(* IEC 61131-3 sources: daoli-st-library/DL_Algo, 207 files *)

(* ---- FB_DL_AdaptiveLeadLag.st ---- *)
(*==============================================================================
 * 组件名称 (Component)  : FB_DL_AdaptiveLeadLag
 * 所属子库 (Sublibrary) : DL_Algo
 * 当前版本 (Version)    : 1.0.0
 * 兼容性   (Platform)   : CODESYS 3.5+ / TwinCAT 3 / 汇川 InoProShop / 施耐德 Machine Expert
 *                         仅依赖 Standard.library（R_TRIG / ABS），零厂商私有库
 * 功能描述 (Function)   : 自适应超前-滞后补偿（误差驱动参数缓调 + 无扰切换）。
 *                         ① 补偿本体：连续式 G(s) = (1 + Tlead·s) / (1 + Tlag·s) 的离散实现
 *                            超前段：yLead = x + Tlead·(x − xPrev) / fDtS
 *                            滞后段：y     = y + (yLead − y) · fDtS / (Tlag + fDtS)
 *                            两段都用 fDtS（调用方给的采样周期，秒），**不做 TIME→数值转换**。
 *                         ② 参数缓调：Tlead 按误差幅值缓升缓降（相位裕度需求随误差增大），
 *                            每拍步长 = fAdaptGain·|fErr|·fDtS，并被 fAdaptRate·fDtS 限幅
 *                            （限幅保证"缓"：参数变化速度受控，不会一拍跳变引起输出突跳）。
 *                            Tlead 始终钳在 [fTleadMin, fTleadMax]。
 *                         ③ 无扰切换：bEnable 上升沿开始，fBlend 以固定步长 fDtS / fRampSec
 *                            从 0 线性升到 1；输出 = 切换前保持值 + blend·(计算值 − 保持值)。
 *                            **不用 TON 的 ET 做斜坡**，因而无 TIME→数值转换（跨平台一致），
 *                            且斜坡长度由 fRampSec 显式给出，可预测、可复现。
 * 接口     (Interface)  : 输入 fIn 输入信号、fErr 跟踪误差（驱动自适应）、fDtS 采样周期（秒）、
 *                         fTleadInit / fTlagInit 初值、fTleadMin / fTleadMax 超前时间限、
 *                         fAdaptGain 自适应增益、fAdaptRate 参数变化率限、fRampSec 无扰斜坡时长、
 *                         fOutMax 输出饱和限、bEnable 使能、bReset 复位；输出 fOut 补偿输出、
 *                         fTleadUsed / fTlagUsed 实际使用参数、fBlend 切换斜坡进度、bActive 已生效、
 *                         bLimited 输出饱和、eState / eCause / bError。
 * 边界     (Boundary)   : ① **属主边界（写死）：本件是补偿器本体，输出 fOut 供上层注入，
 *                         不直接写轴指令/不进闭环回路**；本件不做参数辨识（辨识属 `FB_DL_RlsEstimator`），
 *                         只按误差缓调。
 *                         ② 组态闸：fDtS <= DL_ALL_EPS（除零 + 步长退化）、fTlagInit < 0.0、
 *                         fTleadMin < 0.0、fTleadMax <= fTleadMin、fAdaptGain < 0.0、
 *                         fAdaptRate <= 0.0、fRampSec <= DL_ALL_EPS、fOutMax <= 0.0、任一 NaN
 *                         → 故障锁存，fOut 置 0（安全侧）。
 *                         ③ bEnable=FALSE 语义（R191 声明）：fOut 立即置 0（补偿器禁用即不注入），
 *                         但**保留 fTleadUsed 与内部滞后状态**，下次使能由 fBlend 斜坡重新接续，
 *                         属"冻结参数、清零输出"，与"复位"（参数回初值）不同。
 *                         ④ 单枚 R_TRIG（bReset 与 bEnable 各一枚）段 0 无条件周期刷新。
 *                         ⑤ 故障相迁出唯一路径 = bReset 上升沿（R228B）。
 *                         ⑥ 零全局耦合（无 GVL / 无 VAR_EXTERNAL / 无物理地址）。
 * 分工声明 (Scope)      : 与 `FB_DL_StribeckFrictionComp`（摩擦模型本体）分工——本件是线性
 *                         超前滞后相位补偿，那件是非线性摩擦补偿；两者可并行相加注入，
 *                         但都不自己注入（注入点唯一）。
 * 来源标签 (Source Tag) : T2-1 ◐（公开经典超前-滞后补偿结构与自适应步长思想，参考参数域，
 *                         零代码行复制；固定步长无扰斜坡为本库自研包装）
 * 解除式   (Release)    : bReset 上升沿 ∧ 组态合法 → 清故障、参数回初值、清滞后状态与斜坡。
 *                         自证可满足：复位不依赖锁存量。
 * 码表     (Codes)      : 本件不占用任何全局数字码位。出口为 REAL + BOOL（bActive / bLimited /
 *                         bError）+ ENUM（eState / eCause）；数字码位待主控收口阶段统一派号。
 * 红线自检 (Redline)    : R1 ✓ 零 GVL/VAR_EXTERNAL ｜ R2 ✓ 零 %I/%Q/%M ｜ R3 ✓ 纯 IEC 61131-3
 *                         R4 ✓ 除零闸 + 参数区间闸 + 输出饱和 + NaN 闸 ｜ R5 ✓ 声明逐行同行双语注释
 *                         R6 ✓ ENUM+CASE 含 ELSE ｜ R7 ✓ R_TRIG 段 0 无条件刷新
 * 修订历史 (Revision)   : 2026-11-19  v1.0.0  R46 首版（批次 4 · 序号 17）
 *==============================================================================*)

TYPE E_DL_AllState :
(
    eIdle  := 0,    // 未使能或未完成切换斜坡 / Disabled, ramp not started
    eRamp  := 10,   // 无扰切换斜坡进行中 / Bumpless transfer ramp in progress
    eRun   := 20,   // 补偿器全效运行 / Compensator fully engaged
    eFault := 90    // 组态故障相 / Configuration fault phase
);
END_TYPE

TYPE E_DL_AllCause :
(
    eNone       := 0,   // 无异常 / No anomaly
    eCfgIllegal := 1,   // 组态非法（采样周期/时间限/增益/非有限） / Illegal configuration
    eOutSat     := 2,   // 输出触饱和（补偿量需求超限） / Output saturated
    ePhaseBad   := 3    // 非法相位兜底 / Illegal phase fallback
);
END_TYPE

FUNCTION_BLOCK FB_DL_AdaptiveLeadLag
VAR_INPUT
    fIn        : REAL := 0.0;       // 输入信号 [工程单位] / Input signal [unit]
    fErr       : REAL := 0.0;       // 跟踪误差（驱动自适应） [工程单位] / Tracking error driving the adaptation [unit]
    fDtS       : REAL := 0.001;     // 采样周期，域 > DL_ALL_EPS [s] / Sample period, domain > epsilon [s]
    fTleadInit : REAL := 0.05;      // 超前时间初值，域 >= 0.0 [s] / Initial lead time, >= 0.0 [s]
    fTlagInit  : REAL := 0.20;      // 滞后时间初值，域 >= 0.0 [s] / Initial lag time, >= 0.0 [s]
    fTleadMin  : REAL := 0.01;      // 超前时间下限，域 >= 0.0 [s] / Lead time lower bound, >= 0.0 [s]
    fTleadMax  : REAL := 0.50;      // 超前时间上限，域 > fTleadMin [s] / Lead time upper bound, > lower [s]
    fAdaptGain : REAL := 0.10;      // 自适应增益，域 >= 0.0 [1/s] / Adaptation gain, >= 0.0 [1/s]
    fAdaptRate : REAL := 0.50;      // 参数变化率限，域 > 0.0 [s/s] / Parameter rate limit, > 0.0 [s/s]
    fRampSec   : REAL := 0.20;      // 无扰斜坡时长，域 > DL_ALL_EPS [s] / Bumpless ramp duration, > epsilon [s]
    fOutMax    : REAL := 100.0;     // 输出饱和限，域 > 0.0 [工程单位] / Output saturation limit, > 0.0 [unit]
    bEnable    : BOOL := FALSE;     // 使能；FALSE 时输出置 0 但保留参数 [-] / Enable; FALSE zeroes the output but keeps parameters
    bReset     : BOOL := FALSE;     // 复位，上升沿清故障并使参数回初值 [-] / Reset, clears the fault and restores initial parameters
END_VAR
VAR_OUTPUT
    fOut       : REAL;              // 补偿输出（已饱和） [工程单位] / Compensation output, saturated [unit]
    fTleadUsed : REAL;              // 实际使用中的超前时间 [s] / Lead time in use [s]
    fTlagUsed  : REAL;              // 实际使用中的滞后时间 [s] / Lag time in use [s]
    fBlend     : REAL;              // 切换斜坡进度，域 0..1 [-] / Ramp progress in 0..1
    bActive    : BOOL;              // 补偿器全效生效（blend 已达 1） [-] / Compensator fully engaged
    bLimited   : BOOL;              // 本拍输出触饱和 [-] / Output saturated this scan
    eState     : E_DL_AllState;     // 状态出口 [-] / State outlet
    eCause     : E_DL_AllCause;     // 成因出口（R190 归因唯一） [-] / Cause outlet
    bError     : BOOL;              // 故障标志（组态非法） [-] / Error flag, illegal configuration
END_VAR
VAR
    _eState  : E_DL_AllState := E_DL_AllState.eIdle;    // 内部相位（CASE 唯一写入目标） / Internal phase
    _eCause  : E_DL_AllCause := E_DL_AllCause.eNone;    // 成因出口暂存 / Cause staging
    rtReset  : R_TRIG;              // 复位沿实例，段 0 无条件调用 / Reset edge instance
    rtEnable : R_TRIG;              // 使能沿实例，段 0 无条件调用 / Enable edge instance
    _fTlead  : REAL;                // 超前时间（锁存量） [s] / Lead time, latched [s]
    _fXPrev  : REAL;                // 上拍输入快照（锁存量） [工程单位] / Previous input, latched [unit]
    _fYState : REAL;                // 滞后段内部状态（锁存量） [工程单位] / Lag stage internal state, latched [unit]
    _fBlend  : REAL;                // 斜坡进度（锁存量） [-] / Ramp progress, latched
    _fHold   : REAL;                // 切换前保持值（锁存量） [工程单位] / Value held before transfer, latched [unit]
    _fLead   : REAL;                // 超前段输出当拍量 [工程单位] / Lead-stage output this scan [unit]
    _fComp   : REAL;                // 补偿计算值当拍量 [工程单位] / Computed compensation this scan [unit]
    _fStep   : REAL;                // 参数调整步长当拍量 [s] / Parameter step this scan [s]
    _fRate   : REAL;                // 每拍允许的最大参数变化量 [s] / Maximum parameter change per scan [s]
    _bFault  : BOOL;                // 组态故障锁存位（锁存量） / Latched configuration fault
    _bCfgBad : BOOL;                // 组态非法当拍量 [-] / Illegal configuration this scan
    _bNonFin : BOOL;                // 输入非有限当拍量 [-] / Non-finite input this scan
    _bSat    : BOOL;                // 本拍输出饱和当拍量 [-] / Output saturation this scan
END_VAR
VAR CONSTANT
    DL_ALL_EPS  : REAL := 1.0E-9;   // 时间判零容差（秒级，需比通用 eps 更紧） [无量纲] / Time epsilon in seconds, tighter than usual
    DL_ALL_ONE  : REAL := 1.0;      // 斜坡进度上限 1.0 [无量纲] / Ramp ceiling
    DL_ALL_ZERO : REAL := 0.0;      // 零基准 [无量纲] / Zero baseline
END_VAR

(* —— 段 0：判据派生 + 两沿实例无条件周期刷新 —— *)
_bNonFin := (fIn <> fIn) OR (fErr <> fErr) OR (fDtS <> fDtS)              // NaN 自反判（判等禁令唯一例外） / NaN self-reflexive tests
         OR (fTleadInit <> fTleadInit) OR (fTlagInit <> fTlagInit)
         OR (fTleadMin <> fTleadMin) OR (fTleadMax <> fTleadMax)
         OR (fAdaptGain <> fAdaptGain) OR (fAdaptRate <> fAdaptRate)
         OR (fRampSec <> fRampSec) OR (fOutMax <> fOutMax);
_bCfgBad := (fDtS <= DL_ALL_EPS)                                          // 采样周期闸（除零 + 步长退化） / Sample period gate
         OR (fTleadInit < 0.0) OR (fTlagInit < 0.0)                       // 时间初值非负闸 / Non-negative initial times
         OR (fTleadMin < 0.0) OR (fTleadMax <= fTleadMin)                 // 超前限区间闸 / Lead bounds interval gate
         OR (fAdaptGain < 0.0) OR (fAdaptRate <= 0.0)                     // 自适应增益与速率闸 / Adaptation gain and rate gates
         OR (fRampSec <= DL_ALL_EPS) OR (fOutMax <= 0.0) OR _bNonFin;     // 斜坡与饱和限 + 非有限 / Ramp, saturation limit, non-finite
rtReset(CLK := bReset);                                                   // 复位沿，每拍必调（R228A） / Reset edge, every scan
rtEnable(CLK := bEnable);                                                 // 使能沿，每拍必调 / Enable edge, every scan

(* —— 段 1：单拍量预清零（锁存量 _fTlead/_fXPrev/_fYState/_fBlend/_fHold/_bFault 不入清单） —— *)
fOut     := 0.0;        // 输出每拍预清 / Output preset
fBlend   := 0.0;        // 斜坡出口预清 / Ramp outlet preset
bActive  := FALSE;      // 生效位预清 / Active preset
bLimited := FALSE;      // 饱和位预清 / Limited preset
bError   := FALSE;      // 故障标志预清（R45 配对） / Error flag preset
_bSat    := FALSE;      // 饱和当拍量预清 / Saturation preset

(* —— 段 2：复位沿（参数回初值、清滞后状态与斜坡） —— *)
IF rtReset.Q THEN
    _bFault  := FALSE;                       // 清故障锁存 / Clear the fault latch
    _eCause  := E_DL_AllCause.eNone;         // 清成因 / Clear cause
    _fTlead  := fTleadInit;                  // 超前时间回初值 / Lead time back to the initial value
    _fYState := 0.0;                         // 滞后段状态清零 / Lag state cleared
    _fXPrev  := fIn;                         // 输入快照对齐当拍（防复位首拍伪微分） / Align the snapshot to the present input
    _fBlend  := 0.0;                         // 斜坡清零 / Ramp cleared
    _fHold   := 0.0;                         // 保持值清零 / Hold cleared
    IF _eState = E_DL_AllState.eFault THEN
        _eState := E_DL_AllState.eIdle;      // 故障相迁出（R228B） / Leave fault phase
    END_IF
END_IF
IF _bCfgBad THEN
    _bFault := TRUE;                         // 组态非法锁存 / Latch illegal configuration
    _eCause := E_DL_AllCause.eCfgIllegal;    // 归因：组态非法 / Cause: illegal configuration
END_IF

(* —— 段 3：无扰切换斜坡管理（使能沿起坡；固定步长，无 TIME→数值转换） —— *)
IF rtEnable.Q THEN
    _fHold  := fOut;                         // 记录切换前输出为保持值（若无历史则为 0） / Capture the pre-transfer output
    _fBlend := 0.0;                          // 从 0 起坡 / Start the ramp at zero
    _eState := E_DL_AllState.eRamp;          // 入斜坡相 / Enter the ramp phase
END_IF
IF bEnable AND (NOT _bCfgBad) THEN
    IF _fBlend < DL_ALL_ONE THEN
        _fBlend := _fBlend + (fDtS / fRampSec);     // 固定步长推进（分母已闸） / Fixed-step advance, denominator gated
        IF _fBlend >= DL_ALL_ONE THEN
            _fBlend := DL_ALL_ONE;                  // 上限钳 / Ceiling clamp
            _eState := E_DL_AllState.eRun;           // 斜坡完成，全效运行 / Ramp done, fully engaged
        ELSE
            _eState := E_DL_AllState.eRamp;          // 仍在斜坡 / Still ramping
        END_IF
    END_IF
ELSIF NOT bEnable THEN
    _fBlend := 0.0;                                 // 禁用即清坡（下次使能重新无扰起坡） / Disable clears the ramp
END_IF

(* —— 段 4：自适应参数缓调（误差驱动，速率限幅，区间钳位） —— *)
IF bEnable AND (NOT _bCfgBad) THEN
    _fStep := fAdaptGain * ABS(fErr) * fDtS;                    // 误差驱动的期望步长 [s] / Desired step from the error
    _fRate := fAdaptRate * fDtS;                                // 每拍允许的最大变化量 [s] / Allowed change per scan
    IF _fStep > _fRate THEN
        _fStep := _fRate;                                       // 速率限幅（"缓"调的实现点） / Rate limit, where "slow" is enforced
    END_IF
    IF fErr > 0.0 THEN
        _fTlead := _fTlead + _fStep;                            // 误差为正：加大超前 / Positive error increases the lead
    ELSE
        _fTlead := _fTlead - _fStep;                            // 误差为负：减小超前 / Negative error reduces the lead
    END_IF
    IF _fTlead > fTleadMax THEN
        _fTlead := fTleadMax;                                   // 上限钳 / Upper clamp
    END_IF
    IF _fTlead < fTleadMin THEN
        _fTlead := fTleadMin;                                   // 下限钳 / Lower clamp
    END_IF
END_IF

(* —— 段 5：补偿本体计算（超前段 → 滞后段） —— *)
IF bEnable AND (NOT _bCfgBad) THEN
    _fLead := fIn + (_fTlead * ((fIn - _fXPrev) / fDtS));       // 超前段（分母已闸） / Lead stage, denominator gated
    IF (fTlagInit + fDtS) > DL_ALL_EPS THEN
        _fYState := _fYState + ((_fLead - _fYState) * (fDtS / (fTlagInit + fDtS)));   // 滞后段一阶离散 / Lag stage, first order
    ELSE
        _fYState := _fLead;                                     // 滞后时间为 0 且 dt 病态：直通 / Degenerate case: pass through
    END_IF
    _fComp := _fYState;                                         // 补偿计算值 / Computed compensation
    fOut   := _fHold + (_fBlend * (_fComp - _fHold));           // 无扰混合输出 / Bumpless blended output
    IF fOut > fOutMax THEN
        fOut   := fOutMax;                                      // 正饱和 / Saturate high
        _bSat  := TRUE;
    ELSIF fOut < -fOutMax THEN
        fOut   := -fOutMax;                                     // 负饱和 / Saturate low
        _bSat  := TRUE;
    END_IF
    _fXPrev := fIn;                                             // 输入快照更新（本拍末） / Input snapshot at body end
END_IF

(* —— 段 6：锁存相位迁移闸 —— *)
IF _bFault AND (_eState <> E_DL_AllState.eFault) THEN
    _eState := E_DL_AllState.eFault;                            // 锁存即入故障相 / Latch enters fault phase
END_IF

(* —— 段 7：相位机（ENUM 全成员显式标签 + ELSE 兜底，R128） —— *)
CASE _eState OF

E_DL_AllState.eIdle:
    IF _bFault THEN                                             // 出口 1：组态故障 / Configuration fault
        _eState := E_DL_AllState.eFault;
    ELSIF bEnable THEN                                          // 出口 2：使能到来（无沿也算） / Enable present
        _eState := E_DL_AllState.eRamp;
    END_IF

E_DL_AllState.eRamp:
    IF _bFault THEN                                             // 出口 1：组态故障 / Configuration fault
        _eState := E_DL_AllState.eFault;
    ELSIF (NOT bEnable) THEN                                    // 出口 2：被禁用，回等待相 / Disabled, back to idle
        _eState := E_DL_AllState.eIdle;
    END_IF

E_DL_AllState.eRun:
    IF _bFault THEN                                             // 出口 1：组态故障 / Configuration fault
        _eState := E_DL_AllState.eFault;
    ELSIF NOT bEnable THEN                                      // 出口 2：被禁用，回等待相 / Disabled, back to idle
        _eState := E_DL_AllState.eIdle;
    END_IF

E_DL_AllState.eFault:
    ;                                                           // 故障相：仅段 2 复位沿可迁出 / Only the reset edge leaves this phase

ELSE
    _bFault := TRUE;                                            // 非法相位兜底锁存 / Illegal-phase fallback latch
    _eCause := E_DL_AllCause.ePhaseBad;                         // 归因：非法相位 / Cause: illegal phase
    _eState := E_DL_AllState.eFault;                            // 强拉故障相 / Force fault phase

END_CASE

(* —— 段 8：出口单点映射（名实双出口，R191） —— *)
fTleadUsed := _fTlead;                                          // 超前时间出口 / Lead time outlet
fTlagUsed  := fTlagInit;                                        // 滞后时间出口（本件不调整滞后） / Lag time outlet, not adapted
fBlend     := _fBlend;                                          // 斜坡出口 / Ramp outlet
bActive    := (_eState = E_DL_AllState.eRun) AND (NOT _bFault); // 全效 = 运行相且无故障 / Fully engaged
bLimited   := _bSat;                                            // 饱和出口 / Saturation outlet
bError     := _bFault OR _bCfgBad;                              // 故障标志 = 锁存或组态非法 / Error = latch or illegal config
IF _bSat AND (NOT _bFault) THEN
    _eCause := E_DL_AllCause.eOutSat;                           // 提示：输出饱和（信息级） / Notice: output saturated
END_IF
eState := _eState;                                              // 状态出口 / State outlet
eCause := _eCause;                                              // 成因出口 / Cause outlet

END_FUNCTION_BLOCK

(* ---- FB_DL_CrossLimitSelect.st ---- *)
(*==============================================================================
 * 组件名称 (Component)  : FB_DL_CrossLimitSelect
 * 溯源说明 (Provenance): 道莅 clean-room 防御性实现（IEC 61131-3 纯净实现，闭源文档仅借语义，零代码行）
 * 所属子库 (Sublibrary) : DL_Algo / ProcessControl
 * 当前版本 (Version)    : 1.0.0
 * 兼容性   (Platform)   : CODESYS 3.5 / TwinCAT 3 / 汇川 InoProShop / 施耐德
 *                         Machine Expert；纯 IEC 61131-3（第 3 版），仅用
 *                         Standard.library 的 LIMIT / MIN / MAX / ABS
 * 组件分类 (Category)   : 功能块（FUNCTION_BLOCK）· 燃烧双交叉限幅
 * 功能一句话 (Summary)  : 把主控输出分配成空气/燃气两路给定，按「先行侧自由、
 *                         跟随侧受实测流量约束」的双交叉限幅律钳制，输出限幅
 *                         标志与距限幅点余量。
 *
 * 本件存在的意义 (Why this unit exists)
 *   库内 SplitRangeControl 是单输出分程、RatioController 是比值站，都不解
 *   「空燃两侧谁先给」这个燃烧专有语义。双交叉限幅管的是**同拍的选择律**：
 *   升负荷时先行侧先动、跟随侧被实测流量压住；降负荷时反过来。
 *   写成一件的理由是它必须逐拍可复算（验收向量要能独立手算），
 *   与氧量修正（慢时标积分律，见 FB_DL_ExcessAirTrim）不可合并。
 *
 * 依赖收窄 (Dependency narrowing)
 *   DL_Algo 只允许依赖 Standard.library（DL_Algo/VERSION.md 明示不得引用
 *   DL_Base / DL_MathData）。因此本件的限幅用内建 LIMIT、容差比较与死区
 *   判断全部内联等价实现，不调用任何 DL_ 子库件。此处声明留档（R11 先例）。
 *
 * 折算口径 (Scaling rationale —— 必须写清，否则本件不可复算)
 *   主控输出是 [%]，流量是 [Nm3/h]，两者不同量纲，接口未给阀门流量量程。
 *   本件的折算基准是**实测流量本身**：主控 [%] 与实测流量在当前工况下对应，
 *   故「约束侧的允许百分比」= 主控输出 × (允许流量 / 实测流量)。该比值无量纲，
 *   不引入任何隐藏量程参数。实测流量 ≤ DL_FLOW_EPS 时（点火初期或流量计未投用）
 *   没有折算基准，此时**直接放行主控值**并置信息码，绝不拿 0 做除数。
 *
 * 边界安全 (Boundary)
 *   ① fAirFuelRatio <= 0、fLeadMargin < 1.0、或二者非有限 → 故障 2B10，
 *      **双侧给定归零**（安全侧 = 切断燃料，宁可熄火不可爆燃）；
 *   ② 任一流量或主控非有限 → 故障 2B11，**保持末次有效给定**
 *      （切 0 会熄火/爆燃，与「参数非法」的安全方向相反，两条并列写死）；
 *   ③ 限幅生效 → 信息 2B01（空气侧受限）/ 2B02（燃气侧受限）；
 *   ④ 失能 → 回 eIdle，fAirSp 与 fGasSp **逐个显式赋 0**（R72 双路径清零，
 *      不依赖段尾镜像），bLimited / fLimitMargin 同时清零；
 *   ⑤ 除零前置闸先于任何除法：比率闸在段 3、实测流量闸在段 6，两处都在商之前；
 *   ⑥ 本件无复位引脚，故障态在原因消失后自动回 eNormal（本件无台账需保持，
 *      与 FB_DL_PressureReliefMonitor 的锁存台账件语义不同，已留档）；
 *   ⑦ CASE 落 ELSE 置 2B12 并回 eFault（非法状态兜底）。
 *
 * 错误码    : 16#0002_2B01 空气侧限幅生效（跟随侧为空气）——信息级，正常调节
 *             16#0002_2B02 燃气侧限幅生效（跟随侧为燃气）——信息级，正常调节
 *             16#0002_2B10 空燃比或先行裕度非法（含非有限），双侧给定归零——故障级
 *             16#0002_2B11 输入非有限，保持末次有效给定——故障级，不得切 0
 *             16#0002_2B12 状态机落 ELSE 兜底（非法状态）——故障级，回 eFault
 * 码位总账  : 16#0002_2B01 用 / 16#0002_2B02 用 ｜ 16#0002_2B10 用 / 16#0002_2B11 用 / 16#0002_2B12 用
 * 状态机    : E_DL_CrossLimitState（eIdle / eNormal / eAirLimited / eGasLimited / eFault），
 *             CASE 含 ELSE 兜底，ELSE 置 16#0002_2B12 并回 eFault；失能无条件回 eIdle
 * 采样约定  : 每任务周期调用一次，纯代数运算，无定时器、无积分
 * 依赖说明  : 零 DL_ 子库依赖；仅 Standard.library 的 LIMIT / MIN / MAX / ABS
 * 验收向量  : V1 空气先行、主控 60 %、空气 1200 Nm3/h、燃气 100 Nm3/h、比率 10
 *               → 允许燃气 1200/10×1.05 = 126 → 燃气给定 = 60×126/100 = 75.6 → 钳到 60；
 *               不受限，eNormal，bValid = TRUE
 *             V2 同 V1 但燃气实测 130 Nm3/h（超供）→ 燃气给定 = 60×126/130 = 58.15，
 *               bLimited = TRUE，fLimitMargin = 1.85，eErr = 2B02，eGasLimited
 *             V3 fAirFuelRatio = 0 → 双侧给定 0，eErr = 2B10，bError = TRUE，eFault
 *             V4 fLeadMargin = 0.95 → 双侧给定 0，eErr = 2B10（先行裕度主向量）
 *             V5 fAirFlow = NaN → 给定保持上一拍有效值，eErr = 2B11（保持主向量）
 *             V6 bEnable = FALSE → fAirSp = 0 且 fGasSp = 0，bLimited = FALSE，eIdle
 *             V7 燃气先行（bAirLead = FALSE）+ 空气超供 → eErr = 2B01，eAirLimited
 * 红线自检  : 全局变量声明零使用 / 外部变量访问零使用 / 物理地址零使用 ｜ 纯 IEC 61131-3 ｜ 两处除零
 *             前置闸 ｜ 浮点只用容差与大小比较，无判等 ｜ 无循环 ｜ 全变量双语
 *             同行注释 ｜ ENUM + CASE 含 ELSE ｜ 无定时器实例（无刷新项，天然合规）
 *             ｜ 无魔法数
 * 修订历史  : 2026-11-16  v1.0.0  首版入库（R22 · 批 2 · 燃烧保护律）
 *============================================================================*)

(*-----------------------------------------------------------------------------
 * 枚举: E_DL_CrossLimitState（归属本功能块，同文件发布，全库唯一定义）
 * 含义: 交叉限幅的工作相位。0 起步长 10。
 *-----------------------------------------------------------------------------*)
TYPE E_DL_CrossLimitState :
(
    eIdle       := 0,   // 待机：未使能，双侧给定为 0 / Idle, disabled, both setpoints zero
    eNormal     := 10,  // 正常：跟随侧未被压住，两路等于主控 / Normal, the follower is not constrained
    eAirLimited := 20,  // 空气侧受限：燃气先行时空气被压住 / Air limited, gas leads and air is constrained
    eGasLimited := 30,  // 燃气侧受限：空气先行时燃气被压住 / Gas limited, air leads and gas is constrained
    eFault      := 99   // 故障：参数非法或输入非有限 / Fault, illegal parameter or non-finite input
);
END_TYPE

FUNCTION_BLOCK FB_DL_CrossLimitSelect
VAR_INPUT
    fMasterOut     : REAL;                     // 主控输出 [%]，范围 0~100 / master controller output [%], range 0~100
    fAirFlow       : REAL;                     // 实测空气流量 [Nm3/h] / measured air flow [Nm3/h]
    fGasFlow       : REAL;                     // 实测燃气流量 [Nm3/h] / measured gas flow [Nm3/h]
    fAirFuelRatio  : REAL := 10.0;             // 目标空燃比 [Nm3空气/Nm3燃气]，须 > 0 / target air to fuel ratio [Nm3 air per Nm3 gas], must be > 0
    fLeadMargin    : REAL := 1.05;             // 先行裕度 [倍]，须 >= 1.0 / leading margin [ratio], must be >= 1.0
    bAirLead       : BOOL := TRUE;             // TRUE 空气先行 / FALSE 燃气先行 / TRUE air leads, FALSE gas leads
    bEnable        : BOOL;                     // 使能 / enable
END_VAR
VAR_OUTPUT
    fAirSp         : REAL;                     // 空气给定 [%]，范围 0~100 / air setpoint [%], range 0~100
    fGasSp         : REAL;                     // 燃气给定 [%]，范围 0~100 / gas setpoint [%], range 0~100
    bLimited       : BOOL;                     // 跟随侧限幅生效标志 / follower side limiting active flag
    fLimitMargin   : REAL;                     // 距限幅点余量 [%]，未限幅时为 0 / distance to the limiting point [%], zero when unlimited
    eErr           : UDINT;                    // 错误码，0 表示无错 / error code, 0 means no error
    bError         : BOOL;                     // 故障级标志，仅故障级错误置位 / fault-class flag, set only on fault-level codes
    bValid         : BOOL;                     // 输出可用标志 / outputs usable flag
END_VAR
VAR
    _eState        : E_DL_CrossLimitState := E_DL_CrossLimitState.eIdle; // 当前相位 / current phase
    _eCand         : E_DL_CrossLimitState := E_DL_CrossLimitState.eNormal; // 本拍候选相位 / candidate phase of this scan
    _bInit         : BOOL := FALSE;            // 首扫标志，初值 FALSE 取非判定 / first-scan flag, tested negated
    _bParamBad     : BOOL;                     // 参数非法标志 / illegal parameter flag
    _bFiniteBad    : BOOL;                     // 输入非有限标志 / non-finite input flag
    _bIllegal      : BOOL;                     // 非法状态标志 / illegal state flag
    _bLimC         : BOOL;                     // 本拍限幅标志（候选） / limiting flag of this scan
    _fMarginC      : REAL;                     // 本拍余量（候选）[%] / margin of this scan [%]
    _fMasterUse    : REAL;                     // 生效主控输出 [%]，已钳位 / effective master output [%], clamped
    _fAirHeld      : REAL;                     // 空气给定保持量 [%] / held air setpoint [%]
    _fGasHeld      : REAL;                     // 燃气给定保持量 [%] / held gas setpoint [%]
    _fGasAvail     : REAL;                     // 允许燃气流量 [Nm3/h] / allowable gas flow [Nm3/h]
    _fAirNeed      : REAL;                     // 所需空气流量 [Nm3/h] / required air flow [Nm3/h]
    _fAirAllowed   : REAL;                     // 允许空气流量 [Nm3/h] / allowable air flow [Nm3/h]
    _fSpC          : REAL;                     // 受限侧候选给定 [%] / candidate setpoint of the constrained side [%]
    _fAirC         : REAL;                     // 空气候选给定 [%] / candidate air setpoint [%]
    _fGasC         : REAL;                     // 燃气候选给定 [%] / candidate gas setpoint [%]
END_VAR
VAR CONSTANT
    DL_PCT_MIN     : REAL := 0.0;              // 给定下限 [%] / setpoint floor [%]
    DL_PCT_MAX     : REAL := 100.0;            // 给定上限 [%] / setpoint ceiling [%]
    DL_VAL_LIM     : REAL := 1.0E30;           // 有限性判定的绝对值上限 [无量纲] / finiteness ceiling [dimensionless]
    DL_EPS         : REAL := 1.0E-6;           // 浮点比较容差 [%] / float comparison tolerance [%]
    DL_FLOW_EPS    : REAL := 1.0E-6;           // 折算基准流量下限 [Nm3/h] / scaling base flow floor [Nm3/h]
    DL_RATIO_MIN   : REAL := 0.0;              // 空燃比下限 [Nm3/Nm3]，须严格大于 / ratio floor, must be strictly greater
    DL_LEAD_MIN    : REAL := 1.0;              // 先行裕度下限 [倍] / leading margin floor [ratio]
    DL_LEAD_MAX    : REAL := 10.0;             // 先行裕度上限 [倍]，防呆 / leading margin ceiling [ratio], sanity bound
END_VAR

(*------------------------------------------------------------------------------
 * 段 1｜每拍预置（输出在段 8 单点写入，此处不清；保持量不清）
 *      Per-scan presets, outputs and held values are untouched here
 *-----------------------------------------------------------------------------*)
eErr        := 16#0000_0000;                   // 错误码每拍重算 / error code recomputed every scan
bError      := FALSE;                          // 故障标志每拍重算 / fault flag recomputed every scan
bValid      := FALSE;                          // 可用标志每拍重算 / usable flag recomputed every scan
bLimited    := FALSE;                          // 限幅标志每拍重算 / limiting flag recomputed every scan
fLimitMargin := 0.0;                           // 余量每拍重算 [%] / margin recomputed every scan
_bParamBad  := FALSE;                          // 参数非法标志预清零 / parameter flag pre-cleared
_bFiniteBad := FALSE;                          // 非有限标志预清零 / non-finite flag pre-cleared
_bIllegal   := FALSE;                          // 非法状态标志预清零 / illegal state flag pre-cleared
_bLimC      := FALSE;                          // 候选限幅标志预清零 / candidate limiting flag pre-cleared
_fMarginC   := 0.0;                            // 候选余量预清零 [%] / candidate margin pre-cleared
_eCand      := E_DL_CrossLimitState.eNormal;   // 候选相位预置正常 / candidate phase preset to normal

(*------------------------------------------------------------------------------
 * 段 2｜首扫初始化（给定从 0 起：点火前燃气必须为 0）
 *      First-scan initialisation, setpoints start at zero because gas must be zero before ignition
 *-----------------------------------------------------------------------------*)
IF NOT _bInit THEN
    _eState   := E_DL_CrossLimitState.eIdle;   // 相位待机 / phase idle
    _fAirHeld := 0.0;                          // 空气给定保持量 0 [%] / held air setpoint zero
    _fGasHeld := 0.0;                          // 燃气给定保持量 0 [%] / held gas setpoint zero
    _bInit    := TRUE;                         // 首扫只做一次 / the first scan runs once
END_IF

(*------------------------------------------------------------------------------
 * 段 3｜参数闸门与除零前置闸（比率与先行裕度的合法性先于任何除法）
 *      Parameter gate and the pre-division guard, checked before any division
 *-----------------------------------------------------------------------------*)
IF (fAirFuelRatio <> fAirFuelRatio) OR (ABS(fAirFuelRatio) > DL_VAL_LIM)
   OR (fAirFuelRatio <= DL_RATIO_MIN) THEN
    _bParamBad := TRUE;                        // 空燃比非法或非有限 / ratio illegal or non-finite
END_IF
IF (fLeadMargin <> fLeadMargin) OR (ABS(fLeadMargin) > DL_VAL_LIM)
   OR (fLeadMargin < DL_LEAD_MIN) OR (fLeadMargin > DL_LEAD_MAX) THEN
    _bParamBad := TRUE;                        // 先行裕度非法（须 1.0~10.0） / margin illegal, must be 1.0 to 10.0
END_IF

(*------------------------------------------------------------------------------
 * 段 4｜输入有限性闸门（区间判据同时拦 NaN 与 ±Inf，不做浮点判等）
 *      Input finiteness gate, the interval test catches NaN and infinity alike
 *-----------------------------------------------------------------------------*)
IF (fMasterOut < -DL_VAL_LIM) OR (fMasterOut > DL_VAL_LIM) THEN
    _bFiniteBad := TRUE;                       // 主控输出非有限 / master output non-finite
END_IF
IF (fAirFlow < -DL_VAL_LIM) OR (fAirFlow > DL_VAL_LIM) THEN
    _bFiniteBad := TRUE;                       // 空气流量非有限 / air flow non-finite
END_IF
IF (fGasFlow < -DL_VAL_LIM) OR (fGasFlow > DL_VAL_LIM) THEN
    _bFiniteBad := TRUE;                       // 燃气流量非有限 / gas flow non-finite
END_IF

(*------------------------------------------------------------------------------
 * 段 5｜双交叉限幅计算（仅在使能、参数合法、输入有限时更新保持量）
 *      Cross-limiting computation, the hold values are updated only on valid input
 *-----------------------------------------------------------------------------*)
IF bEnable AND (NOT _bParamBad) AND (NOT _bFiniteBad) THEN
    _fMasterUse := LIMIT(DL_PCT_MIN, fMasterOut, DL_PCT_MAX); // 主控钳进 0~100 % / master clamped
    _fAirC := _fMasterUse;                     // 空气侧先按主控直给 [%] / air follows the master by default
    _fGasC := _fMasterUse;                     // 燃气侧先按主控直给 [%] / gas follows the master by default

    IF bAirLead THEN
        (* 空气先行：燃气侧受实测空气约束（允许燃气 = 空气/比率×裕度） *)
        (* Air leads, gas is constrained by the measured air *)
        IF fAirFuelRatio > DL_RATIO_MIN THEN
            _fGasAvail := (fAirFlow / fAirFuelRatio) * fLeadMargin; // 允许燃气流量 [Nm3/h] / allowable gas flow
            IF fGasFlow > DL_FLOW_EPS THEN
                _fSpC := (_fMasterUse * _fGasAvail) / fGasFlow; // 折算为百分比 [%] / scaled to percent
                _fSpC := LIMIT(DL_PCT_MIN, _fSpC, _fMasterUse); // 跟随侧不得超前主控 [%] / the follower never leads the master
                _fGasC := _fSpC;                   // 燃气候选给定 [%] / candidate gas setpoint
                IF (_fMasterUse - _fGasC) > DL_EPS THEN
                    _bLimC    := TRUE;             // 限幅生效 / limiting active
                    _fMarginC := _fMasterUse - _fGasC; // 距限幅点余量 [%] / distance to the limiting point
                    _eCand    := E_DL_CrossLimitState.eGasLimited; // 燃气侧受限 / gas limited
                END_IF
            END_IF
        END_IF
    ELSE
        (* 燃气先行：空气侧受实测燃气约束（所需空气 = 燃气×比率×裕度） *)
        (* Gas leads, air is constrained by the measured gas *)
        _fAirNeed := fGasFlow * fAirFuelRatio;
        _fAirAllowed := _fAirNeed * fLeadMargin; // 允许空气流量 [Nm3/h] / allowable air flow
        IF fAirFlow > DL_FLOW_EPS THEN
            _fSpC := (_fMasterUse * _fAirAllowed) / fAirFlow; // 折算为百分比 [%] / scaled to percent
            _fSpC := LIMIT(DL_PCT_MIN, _fSpC, _fMasterUse); // 跟随侧不得超前主控 [%] / the follower never leads the master
            _fAirC := _fSpC;                       // 空气候选给定 [%] / candidate air setpoint
            IF (_fMasterUse - _fAirC) > DL_EPS THEN
                _bLimC    := TRUE;                 // 限幅生效 / limiting active
                _fMarginC := _fMasterUse - _fAirC; // 距限幅点余量 [%] / distance to the limiting point
                _eCand    := E_DL_CrossLimitState.eAirLimited; // 空气侧受限 / air limited
            END_IF
        END_IF
    END_IF

    _fAirHeld := LIMIT(DL_PCT_MIN, _fAirC, DL_PCT_MAX); // 双侧钳 0~100 % 后入保持量 / clamped then latched
    _fGasHeld := LIMIT(DL_PCT_MIN, _fGasC, DL_PCT_MAX); // 双侧钳 0~100 % 后入保持量 / clamped then latched
END_IF

(*------------------------------------------------------------------------------
 * 段 6｜相位机（只做迁移；给定值写段 7，绝不在 CASE 内赋值输出）
 *      Phase machine, transitions only, outputs are written in segment seven
 *-----------------------------------------------------------------------------*)
CASE _eState OF

    E_DL_CrossLimitState.eIdle:                 // 待机：参数与输入合法且使能即进入工作相
        IF _bParamBad OR _bFiniteBad THEN
            _eState := E_DL_CrossLimitState.eFault; // 原因未消失，转故障 / the cause persists, go to fault
        ELSIF bEnable THEN
            _eState := _eCand;                  // 按计算结果进入工作相 / enter the working phase from the computation
        END_IF

    E_DL_CrossLimitState.eNormal:               // 正常：跟随侧未被压住
        IF NOT bEnable THEN
            _eState := E_DL_CrossLimitState.eIdle; // 失能回待机 / disabled, back to idle
        ELSIF _bParamBad OR _bFiniteBad THEN
            _eState := E_DL_CrossLimitState.eFault; // 转故障 / go to fault
        ELSE
            _eState := _eCand;                  // 跟随本拍计算结果 / follow this scan's computation
        END_IF

    E_DL_CrossLimitState.eAirLimited:           // 空气侧受限
        IF NOT bEnable THEN
            _eState := E_DL_CrossLimitState.eIdle; // 失能回待机 / disabled, back to idle
        ELSIF _bParamBad OR _bFiniteBad THEN
            _eState := E_DL_CrossLimitState.eFault; // 转故障 / go to fault
        ELSE
            _eState := _eCand;                  // 跟随本拍计算结果 / follow this scan's computation
        END_IF

    E_DL_CrossLimitState.eGasLimited:           // 燃气侧受限
        IF NOT bEnable THEN
            _eState := E_DL_CrossLimitState.eIdle; // 失能回待机 / disabled, back to idle
        ELSIF _bParamBad OR _bFiniteBad THEN
            _eState := E_DL_CrossLimitState.eFault; // 转故障 / go to fault
        ELSE
            _eState := _eCand;                  // 跟随本拍计算结果 / follow this scan's computation
        END_IF

    E_DL_CrossLimitState.eFault:                // 故障：原因消失即自动恢复（本件无复位引脚）
        IF NOT bEnable THEN
            _eState := E_DL_CrossLimitState.eIdle; // 失能回待机 / disabled, back to idle
        ELSIF (NOT _bParamBad) AND (NOT _bFiniteBad) THEN
            _eState := _eCand;                  // 原因消失，自动回工作相 / cause cleared, resume automatically
        END_IF

    ELSE
        _bIllegal := TRUE;                      // 标记非法状态 / flag the illegal state
        _eState   := E_DL_CrossLimitState.eFault; // 回故障态 / back to the fault state
END_CASE

(*------------------------------------------------------------------------------
 * 段 7｜输出发布（优先级链：非法 > 失能 > 参数非法 > 非有限 > 正常）
 *      Output publish by a strict priority chain, every branch writes both setpoints
 *-----------------------------------------------------------------------------*)
IF _bIllegal THEN
    fAirSp       := 0.0;                        // 非法状态：空气给定清零 [%] / illegal state, air zeroed
    fGasSp       := 0.0;                        // 非法状态：燃气给定清零 [%] / illegal state, gas zeroed
    bLimited     := FALSE;                      // 限幅标志清零 / limiting flag cleared
    fLimitMargin := 0.0;                        // 余量清零 [%] / margin cleared
    eErr         := 16#0002_2B12;               // 故障级：状态机兜底 / fault: state machine fallback
    bError       := TRUE;                       // 置故障标志 / raise the fault flag
    bValid       := FALSE;                      // 输出不可用 / outputs unusable
ELSIF NOT bEnable THEN
    fAirSp       := 0.0;                        // 失能：空气给定显式清零 [%] / disabled, air explicitly zeroed
    fGasSp       := 0.0;                        // 失能：燃气给定显式清零 [%] / disabled, gas explicitly zeroed
    bLimited     := FALSE;                      // 限幅标志清零 / limiting flag cleared
    fLimitMargin := 0.0;                        // 余量清零 [%] / margin cleared
    bValid       := FALSE;                      // 失能时输出不可用 / unusable while disabled
ELSIF _bParamBad THEN
    fAirSp       := 0.0;                        // 参数非法：空气给定归零 [%] / illegal parameter, air zeroed
    fGasSp       := 0.0;                        // 参数非法：燃气给定归零（切断燃料，安全侧） [%] / gas zeroed, fuel cut, safe side
    bLimited     := FALSE;                      // 限幅标志清零 / limiting flag cleared
    fLimitMargin := 0.0;                        // 余量清零 [%] / margin cleared
    eErr         := 16#0002_2B10;               // 故障级：空燃比或先行裕度非法 / fault: ratio or margin illegal
    bError       := TRUE;                       // 置故障标志 / raise the fault flag
    bValid       := FALSE;                      // 输出不可用 / outputs unusable
ELSIF _bFiniteBad THEN
    fAirSp       := _fAirHeld;                  // 非有限：保持末次有效空气给定 [%] / hold the last valid air setpoint
    fGasSp       := _fGasHeld;                  // 非有限：保持末次有效燃气给定（不得切 0） [%] / hold the last valid gas setpoint, never zeroed
    bLimited     := FALSE;                      // 限幅标志不宣称（本次未计算） / no limiting claim this scan
    fLimitMargin := 0.0;                        // 余量清零 [%] / margin cleared
    eErr         := 16#0002_2B11;               // 故障级：输入非有限 / fault: non-finite input
    bError       := TRUE;                       // 置故障标志 / raise the fault flag
    bValid       := FALSE;                      // 输出不可用 / outputs unusable
ELSE
    fAirSp       := _fAirHeld;                  // 正常：空气给定 [%] / air setpoint
    fGasSp       := _fGasHeld;                  // 正常：燃气给定 [%] / gas setpoint
    bLimited     := _bLimC;                     // 限幅标志 [%] / limiting flag
    fLimitMargin := _fMarginC;                  // 距限幅点余量 [%] / distance to the limiting point
    IF _bLimC THEN
        IF _eCand = E_DL_CrossLimitState.eAirLimited THEN
            eErr := 16#0002_2B01;               // 信息级：空气侧限幅生效 / informational: air side limiting
        ELSE
            eErr := 16#0002_2B02;               // 信息级：燃气侧限幅生效 / informational: gas side limiting
        END_IF
    END_IF
    bValid := TRUE;                             // 输出可用 / outputs usable
END_IF

END_FUNCTION_BLOCK

(* ---- FB_DL_FlowBalanceCheck.st ---- *)
(*==============================================================================
 * 组件名称 (Component)  : FB_DL_FlowBalanceCheck
 * 所属子库 (Sublibrary) : DL_Algo
 * 当前版本 (Version)    : 1.0.0
 * 兼容性   (Platform)   : CODESYS 3.5+ / TwinCAT 3 / 汇川 InoProShop / 施耐德 Machine Expert
 *                         仅依赖 Standard.library（TON / ABS / MAX），零厂商私有库
 * 功能描述 (Function)   : 多路流量累计平衡校验：每 tWindow 窗口期对有效通道
 *                         重算一次总入 ΣaInflow 与总出 ΣaOutflow，失衡率
 *                           fImbalancePct = (Σin − Σout) ÷ max(|Σin|,|Σout|) × 100
 *                         按容差 fTolPct 与告警阈 fWarnPct 分级出口：
 *                           eBalanced（|失衡| <= fTolPct）/
 *                           eWarn（fTolPct < |失衡| <= fWarnPct）/
 *                           eFault（|失衡| > fWarnPct）。
 *                         通道数钳位 1~8；容差 <= 0 冻结判定并置故障码（规格
 *                         指定）；分母基准过小（无流量）判平衡并置信息码。
 * 接口     (Interface)  : 输入 aInflow 8 路流入累计量、aOutflow 8 路流出累计量
 *                         （同工程单位累计口径）、nChanCnt 有效通道数（钳位
 *                         1~8）、fTolPct 平衡容差 [%]、fWarnPct 告警阈 [%]、
 *                         tWindow 重算窗、bReset 复位；输出 fImbalancePct
 *                         失衡率 [%]、eLevel 分级出口（E_DL_FlowLevel）、
 *                         fSumIn/fSumOut 窗口合计透读、eErrCode 错误码、
 *                         bError 故障标志。
 * 边界     (Boundary)   : ① **属主边界（写死）：本件只做累计量平衡判定，不做
 *                         流量测量、不接管泄漏定位**；单路诊断归通道级件。
 *                         ② 窗口自复位 TON（IN := NOT tonWin.Q，R188），窗到
 *                         （F_TRIG 沿）重算一次，窗内判定输出保持（冻结语义
 *                         声明：非结算拍不重算，规格「窗口期重算」口径）。
 *                         ③ 数组钳位：nChanCnt 钳 [1,8]，越界钳位并置信息码
 *                         eChanClamp；求和界宽 = 钳位后通道数，无越界。
 *                         ④ 分母基准 fBase = MAX(|Σin|,|Σout|)，fBase <
 *                         1E-9 判零流量 → 失衡率 0、eLevel=eBalanced、信息码
 *                         eNoFlow（结构性防除零）。
 *                         ⑤ 组态闸：fTolPct <= 0 或 fWarnPct < fTolPct →
 *                         锁存故障，判定冻结（eLevel 保持上次值，故障拍不重算，
 *                         规格指定），解除沿 = bReset 上升沿（R45 配对）。
 *                         ⑥ 非有限判据（R79 双判）：任一有效通道累计非有限 →
 *                         本窗跳过重算，输出保持，信息码 eInputHold。
 *                         ⑦ 零全局耦合（无 GVL / VAR_EXTERNAL / 物理地址）。
 * 分工声明 (Scope)      : 与 `FB_DL_CoolantLoopBal` 分工：冷却回路专用平衡归
 *                         那件、通用累计平衡判据归本件；与 `FB_DL_Integrator`
 *                         分工：积分归那件，本件只读外部累计量。
 * 来源标签 (Source Tag) : 自研线（质量/体积平衡判据为公开守恒定义 clean-room）
 * 码表     (Codes)      : 本件不占用任何全局数字码位。出口为 LREAL 组 +
 *                         ENUM 分级/错误码；数字码位待主控收口阶段统一派号。
 * 红线自检 (Redline)    : R1 ✓ 零 GVL/VAR_EXTERNAL ｜ R2 ✓ 零 %I/%Q/%M ｜ R3 ✓ 纯 IEC 61131-3
 *                         R4 ✓ 分母防除零 + 通道钳位 + 组态锁存 + 非有限跳过
 *                         ｜ R5 ✓ 声明逐行同行双语注释
 *                         R6 N/A（分级枚举非状态机，无 CASE 迁移） ｜ R7 ✓ 一 TON 一 F_TRIG 一 R_TRIG 段 0 无条件刷新
 * 修订历史 (Revision)   : 2026-11-20  v1.0.0  R50 首版（批次 3 · 序号 11）
 * 验收向量 (Acceptance) : ① nChanCnt=1，Σin=100.0，Σout=99.0，fTolPct=0.5，
 *                         fWarnPct=2.0 → 失衡率 (100−99)/100×100 = 1.0%，
 *                         eLevel=eWarn；② Σin=100.0，Σout=100.0 → 0.0%，
 *                         eBalanced；③ fTolPct=0 → 锁存 eCfgBad，判定冻结；
 *                         ④ Σin=0，Σout=0 → 失衡率 0，eNoFlow 信息码。
 *==============================================================================*)

(*-----------------------------------------------------------------------------
 * 枚举: E_DL_FlowLevel（平衡分级出口）
 *----------------------------------------------------------------------------*)
TYPE E_DL_FlowLevel :
(
    eBalanced := 0,   // 平衡（|失衡率| <= fTolPct） / Balanced within tolerance
    eWarn     := 1,   // 告警（容差与告警阈之间） / Warn band
    eFault    := 2    // 失衡超告警阈 / Imbalance beyond warn threshold
);
END_TYPE

(*-----------------------------------------------------------------------------
 * 枚举: E_DL_FbcErr（错误码；信息级不置 bError，故障级恒伴 bError=TRUE）
 *----------------------------------------------------------------------------*)
TYPE E_DL_FbcErr :
(
    eOk        := 0,   // 正常 / Normal
    eCfgBad    := 1,   // 故障级：容差/告警阈组态非法（判定冻结） / Fault: tolerance config illegal, verdict frozen
    eChanClamp := 2,   // 信息级：通道数越界已钳位 [1,8] / Info: channel count clamped
    eNoFlow    := 3,   // 信息级：窗口合计趋零，按平衡处理 / Info: near-zero flow, deemed balanced
    eInputHold := 4    // 信息级：有效通道含非有限累计，本窗跳过 / Info: non-finite total skipped this window
);
END_TYPE

FUNCTION_BLOCK FB_DL_FlowBalanceCheck
VAR_INPUT
    aInflow  : ARRAY[0..7] OF LREAL;   // 8 路流入累计量（累计口径一致） [工程单位] / Eight inflow totals
    aOutflow : ARRAY[0..7] OF LREAL;   // 8 路流出累计量 [工程单位] / Eight outflow totals
    nChanCnt : UDINT := 8;             // 有效通道数，域 [1,8]（越界钳位） [路] / Active channel count
    fTolPct  : LREAL := 0.5;           // 平衡容差（<=0 故障），域 > 0 [%] / Balance tolerance
    fWarnPct : LREAL := 2.0;           // 告警阈（>= 容差），域 >= fTolPct [%] / Warn threshold
    tWindow  : TIME := T#10S;          // 重算窗时长，域 > T#0S [ms] / Recalculation window
    bReset   : BOOL := FALSE;          // 复位，上升沿清组态锁存 [-] / Reset, rising edge clears cfg latch
END_VAR
VAR_OUTPUT
    fImbalancePct : LREAL;             // 失衡率（窗口结算值，窗间保持） [%] / Imbalance percentage
    eLevel        : E_DL_FlowLevel;    // 分级出口（窗间保持） [-] / Graded verdict outlet
    fSumIn        : LREAL;             // 窗口流入合计透读 [工程单位] / Window inflow sum readout
    fSumOut       : LREAL;             // 窗口流出合计透读 [工程单位] / Window outflow sum readout
    eErrCode      : E_DL_FbcErr;       // 错误码出口 / Error code outlet
    bError        : BOOL;              // 故障标志（组态锁存） [-] / Error flag, latched
END_VAR
VAR
    _nCount   : DINT;                  // 钳位后有效通道数 [路] / Clamped channel count
    _bClamp   : BOOL;                  // 本拍发生通道钳位 [-] / Channel clamp this scan
    _fSumIn   : LREAL;                 // 流入合计中间量 [工程单位] / Inflow sum intermediate
    _fSumOut  : LREAL;                 // 流出合计中间量 [工程单位] / Outflow sum intermediate
    _fBase    : LREAL;                 // 分母基准 = MAX(|Σin|,|Σout|) [工程单位] / Denominator base
    _fImb     : LREAL;                 // 失衡率中间量 [%] / Imbalance intermediate
    _eLevel   : E_DL_FlowLevel := E_DL_FlowLevel.eBalanced;   // 分级锁存（窗间保持源） / Level latch
    _bNonFin  : BOOL;                  // 有效通道非有限当拍量 [-] / Non-finite total this scan
    _bCfgBad  : BOOL;                  // 组态非法当拍量 [-] / Illegal configuration this scan
    _bErrLatch: BOOL;                  // 组态故障锁存位（解除沿 = bReset 上升沿） / Latched config fault
    i         : DINT;                  // 通道循环索引 / Channel loop index
    rtReset   : R_TRIG;                // 复位沿实例，段 0 无条件调用 / Reset edge instance
    ftWin     : F_TRIG;                // 窗结算沿实例，段 0 无条件调用 / Window settlement F_TRIG
    tonWin    : TON;                   // 自复位重算窗（R188），段 0 无条件调用 / Self-resetting window
END_VAR
VAR CONSTANT
    DL_FBC_NMAX  : DINT  := 8;         // 通道定长上限 [路] / Channel ceiling
    DL_FBC_NMIN  : DINT  := 1;         // 通道数下限 [路] / Channel floor
    DL_FBC_ZERO  : LREAL := 0.0;       // 判零基准 [%] / Zero base
    DL_FBC_FLMIN : LREAL := 1.0E-9;    // 分母基准下限（防除零） [工程单位] / Denominator floor
    DL_FBC_HUND  : LREAL := 100.0;     // 百分比换算基 [%] / Percent scale base
END_VAR

(* —— 段 0：通道钳位 + 组态闸 + 窗口/沿无条件刷新 —— *)
_bClamp := FALSE;                      // 钳位量预清 / Clamp preset
_nCount := UDINT_TO_DINT(nChanCnt);    // 通道数转 DINT / Convert count
IF _nCount > DL_FBC_NMAX THEN
    _nCount := DL_FBC_NMAX;            // 上越界钳 8 / Clamp high
    _bClamp := TRUE;                   // 记钳位 / Mark clamp
END_IF
IF _nCount < DL_FBC_NMIN THEN
    _nCount := DL_FBC_NMIN;            // 下越界钳 1 / Clamp low
    _bClamp := TRUE;                   // 记钳位 / Mark clamp
END_IF
_bCfgBad := (fTolPct <= DL_FBC_ZERO) OR (fWarnPct < fTolPct) OR (tWindow <= T#0S);   // 组态域闸（容差/告警阈/窗） / Configuration gate
rtReset(CLK := bReset);                // 复位沿，每拍必调 / Reset edge, every scan
tonWin(IN := (NOT tonWin.Q) AND (NOT _bErrLatch), PT := tWindow);   // 自复位重算窗（故障期停窗，R188） / Self-reset window
ftWin(CLK := tonWin.Q);                // 窗结算沿，每拍必调 / Settlement edge, every scan

(* —— 段 1：复位沿与组态锁存 —— *)
IF rtReset.Q THEN
    _bErrLatch := FALSE;               // 清组态锁存（R188 声明：解除沿 = bReset 上升沿） / Clear cfg latch
END_IF
IF _bCfgBad AND (NOT _bErrLatch) THEN
    _bErrLatch := TRUE;                // 锁存 / Latch
END_IF

(* —— 段 2：有效通道合计与非有限扫描（每拍执行，结算沿取值） —— *)
_fSumIn := DL_FBC_ZERO;                // 合计起步 0 / Sum start zero
_fSumOut := DL_FBC_ZERO;               // 合计起步 0 / Sum start zero
_bNonFin := FALSE;                     // 非有限量预清 / Non-finite preset
FOR i := 0 TO (_nCount - 1) DO
    IF (aInflow[i] <> aInflow[i]) OR ((aInflow[i] - aInflow[i]) <> DL_FBC_ZERO)
       OR (aOutflow[i] <> aOutflow[i]) OR ((aOutflow[i] - aOutflow[i]) <> DL_FBC_ZERO) THEN
        _bNonFin := TRUE;              // 任一有效通道非有限（R79 双判） / Any non-finite total
    END_IF
    _fSumIn := _fSumIn + aInflow[i];   // 流入逐路累计（非有限不写出口，仅置跳过量） / Sum inflow
    _fSumOut := _fSumOut + aOutflow[i];   // 流出逐路累计 / Sum outflow
END_FOR

(* —— 段 3：窗结算重算（故障期冻结；非有限本窗跳过保持上次结论） —— *)
IF ftWin.Q AND (NOT _bErrLatch) THEN
    IF (NOT _bNonFin)
       AND (_fSumIn = _fSumIn) AND ((_fSumIn - _fSumIn) = DL_FBC_ZERO)
       AND (_fSumOut = _fSumOut) AND ((_fSumOut - _fSumOut) = DL_FBC_ZERO) THEN
        fSumIn := _fSumIn;             // 合计落出口 / Sum outlets
        fSumOut := _fSumOut;           // 合计落出口 / Sum outlets
        _fBase := MAX(ABS(_fSumIn), ABS(_fSumOut));   // 分母基准 / Denominator base
        IF _fBase < DL_FBC_FLMIN THEN
            _fImb := DL_FBC_ZERO;      // 零流量：失衡率按 0（防除零，头注释④） / Zero flow: imbalance zero
            _eLevel := E_DL_FlowLevel.eBalanced;       // 按平衡分级 / Deemed balanced
            eErrCode := E_DL_FbcErr.eNoFlow;           // 信息码（不置 bError） / Info code
        ELSE
            _fImb := (_fSumIn - _fSumOut) / _fBase * DL_FBC_HUND;   // 失衡率（分母已过闸） / Imbalance percent
            IF ABS(_fImb) <= fTolPct THEN
                _eLevel := E_DL_FlowLevel.eBalanced;   // 容差内 / Within tolerance
            ELSIF ABS(_fImb) <= fWarnPct THEN
                _eLevel := E_DL_FlowLevel.eWarn;       // 告警带 / Warn band
            ELSE
                _eLevel := E_DL_FlowLevel.eFault;      // 超告警阈 / Beyond warn
            END_IF
        END_IF
        fImbalancePct := _fImb;        // 失衡率落出口 / Imbalance outlet
    END_IF
    (* 非有限本窗跳过：出口保持上次结算值（规格⑥，不重算不抹除） *)
END_IF

(* —— 段 4：出口单点映射（名实双出口同源，R191） —— *)
eLevel := _eLevel;                     // 分级出口 / Level outlet
IF _bErrLatch THEN
    bError := TRUE;                    // 故障标志（R45 配对） / Error flag
    eErrCode := E_DL_FbcErr.eCfgBad;   // 故障级码 / Fault code
ELSE
    bError := FALSE;                   // 无故障级条件 / No fault
    IF NOT ftWin.Q THEN
        IF _bClamp THEN
            eErrCode := E_DL_FbcErr.eChanClamp;   // 信息级：通道钳位 / Info: clamped
        ELSE
            eErrCode := E_DL_FbcErr.eOk;          // 正常 / Normal
        END_IF
    END_IF
    (* 结算拍错误码由段 3 命中分支（eOk/eNoFlow）保留，此处不覆盖 *)
END_IF

END_FUNCTION_BLOCK

(* ---- FB_DL_FrequencySweepGen.st ---- *)
(*==============================================================================
 * 组件名称 (Component)  : FB_DL_FrequencySweepGen
 * 所属子库 (Sublibrary) : DL_Algo
 * 当前版本 (Version)    : 1.0.0
 * 兼容性   (Platform)   : CODESYS 3.5+ / TwinCAT 3 / 汇川 InoProShop / 施耐德 Machine Expert
 *                         仅依赖 Standard.library（TON / ABS），零厂商私有库
 * 功能描述 (Function)   : 频率往返扫描发生器：从 fStartHz 按升斜率 fRampUpHzS
 *                         扫至 fEndHz，边界驻留 tDwell 后按降斜率 fRampDnHzS
 *                         扫回，循环往复。四态顺控：
 *                           eRampUp → eDwellHi → eRampDn → eDwellLo → eRampUp
 *                         输出 fFreqOutHz 当前频率与 bUpward 方向标志。与定频
 *                         （FB_DL_PulseGenerator 频率域）、波形发生、测频
 *                         （FB_DL_FrequencyMeasure）职责三分离（分工声明）。
 * 接口     (Interface)  : 输入 fStartHz 扫描下限（域 > 0）、fEndHz 扫描上限
 *                         （域 > fStartHz）、fRampUpHzS 升斜率（域 > 0）
 *                         [Hz/s]、fRampDnHzS 降斜率（域 > 0） [Hz/s]、tDwell
 *                         边界驻留（域 > T#0S）、bEnable 使能、bReset 复位；
 *                         输出 fFreqOutHz 当前频率 [Hz]、bUpward 升向标志、
 *                         ePhase 四态相位出口、eErrCode 错误码、bError 故障
 *                         标志。
 * 边界     (Boundary)   : ① **属主边界（写死）：本件只出频率给定值，不产生波形、
 *                         不测频、不做定频脉宽**（三分离，分工声明）。
 *                         ② 四态 CASE + ELSE 兜底（R6）；两驻留 TON 与两沿
 *                         实例段 0 无条件调用（R7）；驻留 TON IN 挂相驻留本身
 *                         （R145：不准叠加业务条件补集）。
 *                         ③ 斜率步长 = 斜率 × fCy，单步上限自钳：步长 > 全程
 *                         带宽时按带宽单步直达边界（防步长过冲来回抖动）。
 *                         ④ 组态闸：fStartHz <= 0、fEndHz <= fStartHz、任一
 *                         斜率 <= 0、tDwell <= T#0S → 锁存故障，输出安全侧
 *                         fStartHz 且方向 FALSE，解除沿 = bReset 上升沿
 *                         （R45 配对）。
 *                         ⑤ 非有限判据（R79 双判）：组态量非有限并入组态闸
 *                         （扫频给定源头件，非有限组态不得下放）。
 *                         ⑥ 零全局耦合（无 GVL / VAR_EXTERNAL / 物理地址）。
 * 分工声明 (Scope)      : 与 `FB_DL_FrequencyGenerator` 分工：定频发生归那件、
 *                         往返扫描归本件；与 `FB_DL_FrequencyMeasure` 分工：
 *                         测频归那件；波形合成（正弦/三角）归信号链其他件，
 *                         本件只给频率标量。
 * 来源标签 (Source Tag) : 自研线（往返斜坡扫描为公开测试激励模式 clean-room）
 * 码表     (Codes)      : 本件不占用任何全局数字码位。出口为 LREAL 频率 +
 *                         BOOL 方向 + ENUM 相位/错误码；数字码位待主控收口
 *                         阶段统一派号。
 * 红线自检 (Redline)    : R1 ✓ 零 GVL/VAR_EXTERNAL ｜ R2 ✓ 零 %I/%Q/%M ｜ R3 ✓ 纯 IEC 61131-3
 *                         R4 ✓ 步长过冲自钳 + 组态锁存 + 非有限入闸 ｜ R5 ✓ 声明逐行同行双语注释
 *                         R6 ✓ 四态 CASE 含 ELSE ｜ R7 ✓ 两 TON 一 R_TRIG 段 0 无条件刷新
 * 修订历史 (Revision)   : 2026-11-20  v1.0.0  R50 首版（批次 3 · 序号 13）
 * 验收向量 (Acceptance) : ① fStart=10, fEnd=20, 斜率 100 Hz/s，fCycle=0.01
 *                         → 单步 +1.0 Hz：10 → 11 → … → 20 共 10 拍达上限
 *                         入 eDwellHi，bUpward=TRUE；② tDwell=T#500MS →
 *                         50 拍驻留后转 eRampDn，bUpward=FALSE；③ 斜率
 *                         2000 Hz/s（步长 20 > 带宽 10）→ 单拍直达 20.0
 *                         （过冲自钳，头注释③）；④ fEndHz <= fStartHz →
 *                         锁存 eCfgBad。
 *==============================================================================*)

(*-----------------------------------------------------------------------------
 * 枚举: E_DL_FsgPhase（扫描相位，全库唯一属主本文件）
 *----------------------------------------------------------------------------*)
TYPE E_DL_FsgPhase :
(
    eIdle    := 0,   // 待机（未使能） / Idle
    eRampUp  := 10,  // 升斜坡相 / Up-ramp phase
    eDwellHi := 20,  // 上限驻留相 / Dwell at ceiling phase
    eRampDn  := 30,  // 降斜坡相 / Down-ramp phase
    eDwellLo := 40,  // 下限驻留相 / Dwell at floor phase
    eFault   := 90   // 故障（等复位） / Fault, awaiting reset
);
END_TYPE

(*-----------------------------------------------------------------------------
 * 枚举: E_DL_FsgErr（错误码；故障级恒伴 bError=TRUE）
 *----------------------------------------------------------------------------*)
TYPE E_DL_FsgErr :
(
    eOk       := 0,   // 正常 / Normal
    eCfgBad   := 1,   // 故障级：组态非法（域/斜率/驻留/非有限） / Fault: illegal configuration
    ePhaseBad := 2    // 故障级：非法相位兜底 / Fault: illegal phase fallback
);
END_TYPE

FUNCTION_BLOCK FB_DL_FrequencySweepGen
VAR_INPUT
    fStartHz   : LREAL := 10.0;       // 扫描下限，域 > 0 [Hz] / Sweep floor frequency
    fEndHz     : LREAL := 20.0;       // 扫描上限，域 > fStartHz [Hz] / Sweep ceiling frequency
    fRampUpHzS : LREAL := 100.0;      // 升斜率，域 > 0 [Hz/s] / Upward slope
    fRampDnHzS : LREAL := 100.0;      // 降斜率，域 > 0 [Hz/s] / Downward slope
    tDwell     : TIME := T#500MS;     // 边界驻留时长，域 > T#0S [ms] / Boundary dwell duration
    fCycle     : LREAL := 0.0;        // 扫描周期（<=0 用缺省） [s] / Scan cycle, default used when <= 0
    bEnable    : BOOL := FALSE;       // 使能（FALSE 回待机并归 fStartHz） [-] / Enable
    bReset     : BOOL := FALSE;       // 复位，上升沿清组态锁存并回待机 [-] / Reset, rising edge clears latch
END_VAR
VAR_OUTPUT
    fFreqOutHz : LREAL;               // 当前频率给定输出 [Hz] / Present frequency output
    bUpward    : BOOL;                // 升向标志（TRUE=升斜坡/上限驻留） [-] / Upward direction flag
    ePhase     : E_DL_FsgPhase;       // 四态相位出口 [-] / Phase outlet
    eErrCode   : E_DL_FsgErr;         // 错误码出口 / Error code outlet
    bError     : BOOL;                // 故障标志（组态锁存） [-] / Error flag, latched
END_VAR
VAR
    _eState   : E_DL_FsgPhase := E_DL_FsgPhase.eIdle;   // 内部相（CASE 唯一写入目标） / Internal phase
    _fFreq    : LREAL := 0.0;         // 频率内部锁存（斜坡源） [Hz] / Frequency internal latch
    _fCy      : LREAL;                // 当拍有效周期 [s] / Effective cycle this scan
    _fStepUp  : LREAL;                // 升向单步上限（过冲自钳后） [Hz] / Upward step ceiling
    _fStepDn  : LREAL;                // 降向单步上限 [Hz] / Downward step ceiling
    _fBand    : LREAL;                // 全程带宽 = fEndHz − fStartHz [Hz] / Full band width
    _bNonFin  : BOOL;                 // 组态非有限当拍量 [-] / Non-finite configuration
    _bCfgBad  : BOOL;                 // 组态非法当拍量 [-] / Illegal configuration
    _bErrLatch: BOOL;                 // 组态故障锁存位（解除沿 = bReset 上升沿） / Latched config fault
    _eCause   : E_DL_FsgErr := E_DL_FsgErr.eOk;   // 故障成因锁存（归因唯一，R190） / Latched fault cause
    rtReset   : R_TRIG;               // 复位沿实例，段 0 无条件调用 / Reset edge instance
    tonDwellHi: TON;                  // 上限驻留 TON，段 0 无条件调用（IN 挂相驻留，R145） / Ceiling dwell TON
    tonDwellLo: TON;                  // 下限驻留 TON，段 0 无条件调用 / Floor dwell TON
END_VAR
VAR CONSTANT
    DL_FSG_CYDEF : LREAL := 0.01;     // 缺省扫描周期 [s] / Default scan cycle
    DL_FSG_ZERO  : LREAL := 0.0;      // 判零基准 [Hz] / Zero base
END_VAR

(* —— 段 0：非有限判 + 组态闸 + 周期派生 + 两 TON 一沿无条件刷新 —— *)
_bNonFin := (fStartHz <> fStartHz) OR ((fStartHz - fStartHz) <> DL_FSG_ZERO)
         OR (fEndHz <> fEndHz) OR ((fEndHz - fEndHz) <> DL_FSG_ZERO)
         OR (fRampUpHzS <> fRampUpHzS) OR ((fRampUpHzS - fRampUpHzS) <> DL_FSG_ZERO)
         OR (fRampDnHzS <> fRampDnHzS) OR ((fRampDnHzS - fRampDnHzS) <> DL_FSG_ZERO);   // 组态非有限（R79 双判） / Non-finite configuration
_bCfgBad := _bNonFin OR (fStartHz <= DL_FSG_ZERO) OR (fEndHz <= fStartHz)
         OR (fRampUpHzS <= DL_FSG_ZERO) OR (fRampDnHzS <= DL_FSG_ZERO)
         OR (tDwell <= T#0S);        // 组态域闸 / Configuration gate
IF fCycle > DL_FSG_ZERO THEN
    _fCy := fCycle;                  // 组态周期有效 / Configured cycle valid
ELSE
    _fCy := DL_FSG_CYDEF;            // 周期缺省兜底 / Default cycle fallback
END_IF
_fBand := fEndHz - fStartHz;         // 带宽（组态闸后恒正） / Band width
_fStepUp := MIN(fRampUpHzS * _fCy, _fBand);   // 升步长过冲自钳（头注释③） / Up step clamped to band
_fStepDn := MIN(fRampDnHzS * _fCy, _fBand);   // 降步长过冲自钳 / Down step clamped
rtReset(CLK := bReset);              // 复位沿，每拍必调 / Reset edge, every scan
tonDwellHi(IN := (_eState = E_DL_FsgPhase.eDwellHi), PT := tDwell);   // 上限驻留计时（相驻留使能，出相自复位） / Ceiling dwell timer
tonDwellLo(IN := (_eState = E_DL_FsgPhase.eDwellLo), PT := tDwell);   // 下限驻留计时 / Floor dwell timer

(* —— 段 1：复位沿与组态锁存 —— *)
IF rtReset.Q THEN
    _bErrLatch := FALSE;             // 清组态锁存（R188 声明：解除沿 = bReset 上升沿） / Clear cfg latch
END_IF
IF _bCfgBad AND (NOT _bErrLatch) THEN
    _bErrLatch := TRUE;              // 锁存 / Latch
    _eCause := E_DL_FsgErr.eCfgBad;  // 归因：组态非法 / Cause: config illegal
END_IF

(* —— 段 2：使能退出 → 待机（先于 CASE，退出语义优先） —— *)
IF (NOT bEnable) OR _bErrLatch THEN
    _eState := E_DL_FsgPhase.eIdle;  // 未使能/故障回待机（R191 声明：频率归 fStartHz 安全值） / Back to idle
    _fFreq := fStartHz;              // 频率安全侧归下限 / Frequency safe-side floor
    bUpward := FALSE;                // 方向安全侧 FALSE / Direction safe side
END_IF

(* —— 段 3：四态顺控（仅使能且无故障期推进） —— *)
IF bEnable AND (NOT _bErrLatch) THEN
    CASE _eState OF

    E_DL_FsgPhase.eIdle:
        _fFreq := fStartHz;          // 起扫频率归下限 / Start at floor
        _eState := E_DL_FsgPhase.eRampUp;   // 使能即入升斜坡 / Enter up-ramp on enable

    E_DL_FsgPhase.eRampUp:
        IF _fFreq + _fStepUp >= fEndHz THEN
            _fFreq := fEndHz;        // 步内到顶：贴上限（禁过冲） / Reach ceiling
            _eState := E_DL_FsgPhase.eDwellHi;   // 入上限驻留 / Enter ceiling dwell
        ELSE
            _fFreq := _fFreq + _fStepUp;   // 升斜坡步进 / Up-ramp step
        END_IF

    E_DL_FsgPhase.eDwellHi:
        IF tonDwellHi.Q THEN
            _eState := E_DL_FsgPhase.eRampDn;   // 驻留到：反向 / Dwell done: reverse
        END_IF

    E_DL_FsgPhase.eRampDn:
        IF _fFreq - _fStepDn <= fStartHz THEN
            _fFreq := fStartHz;      // 步内到底：贴下限 / Reach floor
            _eState := E_DL_FsgPhase.eDwellLo;   // 入下限驻留 / Enter floor dwell
        ELSE
            _fFreq := _fFreq - _fStepDn;   // 降斜坡步进 / Down-ramp step
        END_IF

    E_DL_FsgPhase.eDwellLo:
        IF tonDwellLo.Q THEN
            _eState := E_DL_FsgPhase.eRampUp;   // 驻留到：再升 / Dwell done: ramp up again
        END_IF

    E_DL_FsgPhase.eFault:
        ;                            // 故障相驻留（由段 2 迁出链处理） / Held by exit chain

    ELSE
        _bErrLatch := TRUE;          // 非法相位兜底：锁存（R45 配对见段 5） / Illegal phase fallback latch
        _eCause := E_DL_FsgErr.ePhaseBad;   // 归因：非法相位（独立码，R190） / Cause: illegal phase
        _eState := E_DL_FsgPhase.eFault;   // 强拉故障相 / Force fault phase

    END_CASE
END_IF

(* —— 段 4：出口单点映射（名实双出口同源，R191） —— *)
fFreqOutHz := _fFreq;                // 频率出口 / Frequency outlet
bUpward := (_eState = E_DL_FsgPhase.eRampUp) OR (_eState = E_DL_FsgPhase.eDwellHi);   // 方向标志（相别派生单源） / Direction from phase
ePhase := _eState;                   // 相位出口 / Phase outlet
IF _bErrLatch THEN
    bError := TRUE;                  // 故障标志（R45 配对） / Error flag
    eErrCode := _eCause;             // 成因锁存回放（R189） / Cause replay
ELSE
    bError := FALSE;                 // 无故障级条件 / No fault
    eErrCode := E_DL_FsgErr.eOk;     // 正常码 / OK code
END_IF

END_FUNCTION_BLOCK

(* ---- FB_DL_LoopPerfIndex.st ---- *)
(*==============================================================================
 * 组件名称 (Component)  : FB_DL_LoopPerfIndex
 * 所属子库 (Sublibrary) : DL_Algo
 * 当前版本 (Version)    : 1.0.0
 * 兼容性   (Platform)   : CODESYS 3.5+ / TwinCAT 3 / 汇川 InoProShop / 施耐德 Machine Expert
 *                         仅依赖 Standard.library（TON / R_TRIG / ABS / MIN / MAX）与库内
 *                         TIME 换算内核 FC_DL_TimeToLrealSec，零厂商私有库
 * 功能描述 (Function)   : 回路性能指标采集与评价（只出指标与建议档，**不做自整定**）。
 *                         阶跃发生后开窗采集：IAE（绝对误差积分）、ISE（误差平方积分）、
 *                         超调百分比、衰减比（相邻两峰比）、过零振荡计数（带去抖）。
 *                         相序：eIdle（非自动/未使能）→ eCollect（阶跃后窗口采集）→
 *                         eEval（一次算出全部指标）→ eDone（保持到撤自动）。窗口到点由
 *                         TON 单点置位（wording：窗口到时由 tonWindow.Q 单拍事件驱动）。
 * 分工声明 (Scope)      : 自整定属主为 `FB_DL_RelayAutoTune` / `FB_DL_AutoTuneRelay`；
 *                         本件**只测量、只给建议档**（偏快/合适/偏慢/振荡），不修改任何 PID 参数、
 *                         不输出激励信号。若上层把 eTuneHint 直接写进 PID 即为越权使用。
 * 接口     (Interface)  : 输入 fSp 设定、fPv 测量、bInAuto 自动态、bEnable 使能、fStepMin
 *                         阶跃判别门限、tWindow 采集窗时长、tTaskPeriod 调用任务周期、fSettleBandPct
 *                         入窗判据带、fOscHystPct 过零去抖带、bReset 复位；输出 fIae / fIse /
 *                         fOvershootPct / fDecayRatio / nOscCount 五指标、eTuneHint 建议档、
 *                         bEvalDone 评价完成单拍、eState / eCause / bError / nErrId。
 * 边界     (Boundary)   : ① 阶跃判据用容差（|ΔfSp| > fStepMin），浮点禁判等；
 *                         ② 窗口到时由 TON 单点置位；能量积分用 LREAL 中间量，防 REAL 逐拍
 *                         累积溢出（REAL 只有 24 位有效位，1e7 拍后即饱和）；
 *                         ③ 测量非有限 → 该拍剔除并计数，连续超过 5 拍置故障（单拍毛刺不断线）；
 *                         ④ 组态闸：fStepMin <= 0.0、tWindow <= T#0S、tTaskPeriod <= T#0S、
 *                         fSettleBandPct <= 0.0、fOscHystPct <= 0.0 或任一浮点引脚 NaN → 故障锁存；
 *                         ⑤ TON 一枚 + R_TRIG 一枚段 0 无条件周期刷新；
 *                         ⑥ 故障相迁出唯一路径 = bReset 上升沿；⑦ 零全局耦合（无 GVL / 无物理地址）。
 * 遗留假设 (Assumption) : 【R95 三句声明】① 代理值 = 引脚 tTaskPeriod（调用方任务周期），用于把
 *                         逐拍误差换算成秒；② 覆盖范围 = 任务周期 1 ms ~ 1000 ms 的周期任务与
 *                         自由运行任务的等效周期；③ 覆盖不到的区间（事件任务、抖动 > 50% 的
 *                         超载任务）由调用方负责：这类工况下积分量只作相互比较用，不可与
 *                         示波器实测 IAE 绝对值对拍。该假设已挂入编译验证债。
 * 解除式   (Release)    : bReset 上升沿 ∧ 组态合法 ∧ 非自动态（NOT bInAuto）。
 *                         自证可满足（终审两式 1）：bInAuto 是外部引脚，切手动即可满足；
 *                         该因子**必须是析取语义里的必要条件之一而非恒假组合**——若写成
 *                         「复位沿 ∧ 自动态」则自动态下复位永远清不掉故障（R152 反例），
 *                         本件按「非自动态」实现，解除可达。
 * 码表     (Codes)      : 16#0002_03B2 故障级：回路性能指标故障总码（组态非法 / 测量持续非有限 /
 *                         非法相位），锁存至 bReset 上升沿，归因由 eCause 承载（R190 单件单总码）；
 *                         16#0002_04B5 信息级：本次评价完成（指标已定稿，附建议档）。
 *                         加码反证（R90）：评价完成与「窗口未开」在五指标数值上不可区分
 *                         （未开窗时指标全为上次值或 0），且 bEvalDone 只是单拍位不进台账，
 *                         故须立一码；信息码只在 eEval 迁移那一拍发出。
 *                         码段说明：0002 段故障子带 03xx / 信息子带 04xx，本件取 03B2 / 04B5
 *                         （源码实扫该两槽为空，续接同子带已用最大值，未回填碎片孔洞）。
 * 编译门槛 (Build Gate) : 本件委托 FC_DL_TimeToLrealSec（内部转调平台内建 TIME_TO_LREAL），
 *                         交付门槛：须在 CODESYS / TwinCAT 3 / InoProShop 三平台各编译验证一次。
 * 开源溯源 (Origin)     : 道莅自研 clean-room（参考公开回路性能指标定义与参数域，零代码行复制；
 *                         t2-5-modpid 参数域族）
 * 修订历史 (Revision)   : 2026-11-19  v1.0.0  R45 首版（批次 2 · 序号 8）
 *==============================================================================*)

TYPE E_DL_LpiState :
(
    eIdle    := 0,     // 非自动或未使能，等待阶跃 / Idle, awaiting a setpoint step
    eCollect := 10,    // 窗口采集 / Collecting inside the window
    eEval    := 20,    // 一次求解全部指标 / Evaluating all indices once
    eDone    := 50,    // 评价完成保持 / Done, result held
    eFault   := 90     // 故障锁存相 / Fault latched phase
);
END_TYPE

TYPE E_DL_LpiCause :
(
    eNone        := 0,   // 无故障成因 / No cause
    eCfgIllegal  := 1,   // 组态非法 / Illegal configuration
    eNonFinRun   := 2,   // 测量连续非有限 / Measurement non-finite too long
    ePhaseBad    := 3    // 非法相位兜底 / Illegal phase fallback
);
END_TYPE

TYPE E_DL_LpiHint :
(
    eSuitable   := 0,    // 合适：超调与衰减比均在线内 / Suitable, overshoot and decay ratio within band
    eTooFast    := 10,   // 偏快：超调偏大或衰减比偏大 / Too fast, overshoot or decay ratio high
    eTooSlow    := 20,   // 偏慢：超调过小且响应迟滞 / Too slow, overshoot too small
    eOscillating := 30   // 振荡：过零次数多或衰减比接近 1 / Oscillating, many crossings or decay ratio near one
);
END_TYPE

FUNCTION_BLOCK FB_DL_LoopPerfIndex
VAR_INPUT
    fSp           : REAL := 0.0;        // 设定值 [工程单位] / Setpoint [unit]
    fPv           : REAL := 0.0;        // 测量值 [工程单位] / Process value [unit]
    bInAuto       : BOOL := FALSE;      // 回路在自动态（采集前置条件） [-] / Loop in automatic mode, precondition for collection
    bEnable       : BOOL := TRUE;       // 指标采集使能 [-] / Index collection enable
    fStepMin      : REAL := 1.0;        // 阶跃判别门限，域 > 0.0 [工程单位] / Step detection threshold, domain > 0.0 [unit]
    tWindow       : TIME := T#30S;      // 采集窗时长，域 > T#0S [ms] / Collection window duration, domain > T#0S [ms]
    tTaskPeriod   : TIME := T#10MS;     // 调用任务周期（代理值，见头注释遗留假设），域 > T#0S [ms] / Task period proxy, domain > T#0S [ms]
    fSettleBandPct: REAL := 5.0;        // 入窗判据带（相对阶跃量百分比），域 > 0.0 [%] / Settling band relative to step, domain > 0.0 [%]
    fOscHystPct   : REAL := 1.0;        // 过零去抖带（相对阶跃量百分比），域 > 0.0 [%] / Zero-crossing debounce band, domain > 0.0 [%]
    bReset        : BOOL := FALSE;      // 复位命令，上升沿清故障 [-] / Reset command, rising edge clears fault
END_VAR
VAR_OUTPUT
    fIae          : REAL;               // 绝对误差积分 [工程单位·s] / Integral of absolute error [unit s]
    fIse          : REAL;               // 误差平方积分 [工程单位²·s] / Integral of squared error [unit2 s]
    fOvershootPct : REAL;               // 超调百分比 [%] / Overshoot percentage [%]
    fDecayRatio   : REAL;               // 衰减比（相邻两峰比），0~1 越好 [p.u.] / Decay ratio of adjacent peaks [p.u.]
    nOscCount     : INT;                // 过零振荡计数（已去抖） [次] / Zero-crossing oscillation count, debounced
    eTuneHint     : E_DL_LpiHint;       // 整定建议档（只建议不整定） [-] / Tuning hint, advisory only
    bEvalDone     : BOOL;               // 评价完成单拍位 [-] / Single-scan evaluation done flag
    eState        : E_DL_LpiState;      // 状态出口，段 6 单点映射 / State outlet
    eCause        : E_DL_LpiCause;      // 故障成因出口（R190 归因唯一） / Fault cause outlet
    bError        : BOOL;               // 故障锁存标志 [-] / Fault latch flag
    nErrId        : UDINT;              // 事件码，0 = 无事件 / Event code, 0 = no event
END_VAR
VAR
    _eState       : E_DL_LpiState := E_DL_LpiState.eIdle;   // 内部相位（CASE 唯一写入目标） / Internal phase
    _eCause       : E_DL_LpiCause := E_DL_LpiCause.eNone;   // 故障成因锁存（锁存量） / Latched cause
    tonWindow     : TON;                // 采集窗计时，段 0 无条件调用 / Collection window timer
    rtReset       : R_TRIG;             // 复位沿实例，段 0 无条件调用 / Reset edge
    _fTsSec       : LREAL;              // 任务周期秒数（当拍量） [s] / Task period in seconds
    _uConvErr     : UDINT;              // 时间换算内核错误码（当拍量） [-] / Time-conversion kernel error code
    _bConvErr     : BOOL;               // 时间换算内核故障位（当拍量） [-] / Time-conversion kernel fault flag
    _bConvValid   : BOOL;               // 时间换算内核有效位（当拍量） [-] / Time-conversion kernel valid flag
    _fIaeAcc      : LREAL;              // IAE 累加器（LREAL 防溢出，锁存量） [工程单位·s] / IAE accumulator in LREAL, latched
    _fIseAcc      : LREAL;              // ISE 累加器（LREAL 防溢出，锁存量） [工程单位²·s] / ISE accumulator in LREAL, latched
    _fErr         : REAL;               // 本拍误差 [工程单位] / Error this scan
    _fStepAmp     : REAL;               // 本次阶跃幅值（带符号） [工程单位] / Step amplitude with sign
    _fPvPeak      : REAL;               // 峰值跟踪（锁存量，入窗后开始累积） [工程单位] / Peak tracking, latched, armed after entering band
    _bBandArmed   : BOOL;               // 峰值累积武装位（首次入窗后置位，锁存量） [-] / Peak accumulation armed after first band entry
    _fPeakLast    : REAL;               // 最近一次过零前峰值偏差（锁存量） [工程单位] / Latest pre-crossing peak deviation
    _fPeakPrev    : REAL;               // 上一次过零前峰值偏差（锁存量） [工程单位] / Previous pre-crossing peak deviation
    _fCrossRef    : REAL;               // 过零参考电平（锁存量） [工程单位] / Crossing reference level, latched
    _bCrossSign   : BOOL;               // 上个去抖后误差符号（锁存量） [-] / Debounced error sign, latched
    _nOscAcc      : INT;                // 振荡累计（锁存量） [次] / Oscillation count accumulator, latched
    _nNonFinRun   : INT;                // 非有限连续计数（锁存量） [拍] / Consecutive non-finite scans, latched
    _fSpPrev      : REAL;               // 上拍设定快照（锁存量） [工程单位] / Previous-scan setpoint snapshot
    _fRatios      : REAL;               // 衰减比中间量 [p.u.] / Decay ratio intermediate
    _bNonFin      : BOOL;               // 本拍测量非有限 [-] / Non-finite measurement this scan
    _bCfgBad      : BOOL;               // 组态非法当拍量 [-] / Illegal configuration
    _bStep        : BOOL;               // 阶跃发生当拍量 [-] / Step detected this scan
    _bFault       : BOOL;               // 故障锁存位（锁存量） / Latched fault bit
    _uFault       : UDINT;              // 故障码锁存（锁存量） / Latched fault code
    _uInfo        : UDINT;              // 信息码，每拍重算 / Info code, recomputed each scan
END_VAR
VAR CONSTANT
    DL_FLOAT_EPS  : REAL := 1.0E-6;     // 浮点判零容差（除子统一口径） [无量纲] / Float epsilon for zero tests
    DL_NONFIN_MAX : INT := 5;           // 非有限连续拍数上限（超限置故障） [拍] / Consecutive non-finite limit [scan]
END_VAR

(* —— 段 0：当拍判据派生 + 定时器与沿实例无条件周期刷新 —— *)
_fTsSec := FC_DL_TimeToLrealSec(tIn := tTaskPeriod, eErr => _uConvErr, bError => _bConvErr, bValid => _bConvValid);   // 委托时间换算内核取秒数（R140 委托优先） / Delegate to time kernel for seconds
_bNonFin  := (fSp <> fSp) OR (fPv <> fPv);                                                      // NaN 自反判（判等禁令唯一例外） / NaN self-reflexive tests
_bCfgBad  := (fStepMin <= 0.0) OR (tWindow <= T#0S) OR (tTaskPeriod <= T#0S)                    // 组态域闸（R151 全覆盖） / Config gate
             OR (fSettleBandPct <= 0.0) OR (fOscHystPct <= 0.0)                                 // 判据带正域闸 / Band gates
             OR (fStepMin <> fStepMin) OR (fSettleBandPct <> fSettleBandPct)                     // 参数 NaN 判 / Parameter NaN tests
             OR (fOscHystPct <> fOscHystPct) OR (_uConvErr <> 16#0000_0000);                     // 换算错误并入组态闸 / Conversion error folded into config gate
_bStep := ABS(fSp - _fSpPrev) > fStepMin;                                                        // 阶跃判据（容差式，禁判等） / Step criterion, tolerance-based
rtReset(CLK := bReset);                                                                          // 复位沿，每拍必调（R228A） / Reset edge
tonWindow(IN := (_eState = E_DL_LpiState.eCollect), PT := tWindow);                              // 采集窗计时，IN 由相位派生 / Window timer, IN from phase

(* —— 段 1：单拍量预清零（锁存量与快照量不入清单，R107） —— *)
_uInfo      := 16#0000_0000;       // 信息码每拍重算 / Info recomputed every scan
bEvalDone   := FALSE;              // 完成单拍位每拍预清，唯一分支置位（R44 范式） / Done flag preset
nErrId      := 16#0000_0000;       // 事件码缺省无事件 / Event code default none
bError      := FALSE;              // 故障标志每拍预清，故障分支同拍置位（R45 配对） / Flag preset

(* —— 段 2：复位沿 + 组态域闸 + 连续非有限计数 —— *)
IF rtReset.Q THEN                                                        // 当拍复位沿 / current-scan reset edge
    _bFault := FALSE;                                                    // 清故障锁存位（锁存量） / Clear fault latch
    _uFault := 16#0000_0000;                                             // 清故障锁存码（锁存量） / Clear latched code
    _eCause := E_DL_LpiCause.eNone;                                      // 清成因（锁存量） / Clear latched cause
    IF _eState = E_DL_LpiState.eFault THEN
        _eState := E_DL_LpiState.eIdle;                                  // 故障相迁出唯一路径 / Sole exit from fault phase
    END_IF
END_IF
IF _bCfgBad THEN                                                         // 组态域闸 / Configuration gate
    _uFault := 16#0002_03B2;                                             // 故障级：回路性能指标故障总码 / Fault-level: index fault code
    _bFault := TRUE;
    bError  := TRUE;                                                     // 故障标志同拍置位（R45 配对） / Error flag set same scan
    _eCause := E_DL_LpiCause.eCfgIllegal;                                // 归因：组态非法 / Cause: illegal configuration
END_IF
IF _bNonFin THEN                                                         // 测量非有限：该拍剔除并计数 / Non-finite measurement, drop and count
    IF _nNonFinRun < DL_NONFIN_MAX THEN
        _nNonFinRun := _nNonFinRun + 1;
    END_IF
ELSE
    _nNonFinRun := 0;                                                    // 恢复有限即清连续计数 / Reset counter on finite value
END_IF
IF (NOT _bFault) AND (_nNonFinRun >= DL_NONFIN_MAX) THEN                 // 连续越限置故障 / Consecutive overrun
    _uFault := 16#0002_03B2;
    _bFault := TRUE;
    bError  := TRUE;
    _eCause := E_DL_LpiCause.eNonFinRun;                                 // 归因：测量持续非有限 / Cause: sustained non-finite
END_IF

(* —— 段 3：指标采集（仅 eCollect 相且测量有限时累加） —— *)
IF (_eState = E_DL_LpiState.eCollect) AND (NOT _bNonFin) AND (NOT _bFault) THEN
    _fErr := fSp - fPv;                                                  // 本拍误差 / Error this scan
    _fIaeAcc := _fIaeAcc + ABS(_fErr) * _fTsSec;                         // IAE 累加（LREAL） / IAE accumulation
    _fIseAcc := _fIseAcc + _fErr * _fErr * _fTsSec;                      // ISE 累加（LREAL） / ISE accumulation
    IF (NOT _bBandArmed) AND (ABS(_fErr) <= (ABS(_fStepAmp) * fSettleBandPct * 0.01)) THEN   // 首次入窗才武装峰值累积（R144） / Arm peak accumulation on first band entry
        _bBandArmed := TRUE;
        _fPvPeak := fSp;                                                 // 峰值初值取设定量而非回读量（R144） / Peak seeded from setpoint, not from PV
    END_IF
    IF _bBandArmed THEN
        IF _fStepAmp > 0.0 THEN
            IF fPv > _fPvPeak THEN
                _fPvPeak := fPv;                                         // 上行阶跃：跟踪最高测量 / Upward step peak tracking
            END_IF
        ELSE
            IF fPv < _fPvPeak THEN
                _fPvPeak := fPv;                                         // 下行阶跃：跟踪最低测量 / Downward step peak tracking
            END_IF
        END_IF
    END_IF
    IF ABS(_fErr) > (ABS(_fStepAmp) * fOscHystPct * 0.01) THEN           // 去抖：误差需超出滞环带才更新符号 / Debounce before sign update
        IF _bCrossSign AND (_fErr < 0.0) THEN                            // 正 → 负过零 / Positive to negative crossing
            _fPeakPrev := _fPeakLast;                                    // 峰值队列后移 / Shift peak queue
            _fPeakLast := ABS(_fCrossRef);
            _nOscAcc := _nOscAcc + 1;                                    // 振荡计数递增 / Oscillation count increment
            _bCrossSign := FALSE;
        ELSIF (NOT _bCrossSign) AND (_fErr > 0.0) THEN                   // 负 → 正过零 / Negative to positive crossing
            _fPeakPrev := _fPeakLast;
            _fPeakLast := ABS(_fCrossRef);
            _nOscAcc := _nOscAcc + 1;
            _bCrossSign := TRUE;
        END_IF
        _fCrossRef := _fErr;                                             // 过零参考电平更新 / Update crossing reference
    END_IF
END_IF

(* —— 段 4：阶跃检测（进相前置，同时清采集量） —— *)
IF (NOT _bFault) AND bEnable AND bInAuto AND _bStep AND (_eState <> E_DL_LpiState.eCollect) THEN
    _fStepAmp := fSp - _fSpPrev;                                         // 阶跃幅值（带符号） / Step amplitude with sign
    _fIaeAcc := 0.0;                                                     // 采集量唯一重置点 / Sole reset point for accumulators
    _fIseAcc := 0.0;
    _fPvPeak := fSp;                                                     // 峰值初值取设定量 / Peak seeded from setpoint
    _bBandArmed := FALSE;                                                // 峰值累积重新武装 / Re-arm peak accumulation
    _fPeakLast := 0.0;                                                   // 峰值队列清空 / Clear peak queue
    _fPeakPrev := 0.0;
    _fCrossRef := 0.0;
    _bCrossSign := FALSE;
    _nOscAcc := 0;                                                       // 振荡计数清零 / Clear oscillation count
    _eState := E_DL_LpiState.eCollect;                                   // 进采集相 / Enter collection phase
END_IF
_fSpPrev := fSp;                                                         // 设定快照（主体末更新） / Setpoint snapshot at body end

(* —— 段 5：故障解除式（R240 全当拍量；非自动态为可达必要条件） —— *)
IF rtReset.Q AND (NOT _bCfgBad) AND (NOT bInAuto) THEN
    _bFault := FALSE;                                                    // 清故障锁存位（锁存量） / Clear fault latch
    _uFault := 16#0000_0000;                                             // 清故障锁存码（锁存量） / Clear latched code
    _eCause := E_DL_LpiCause.eNone;                                      // 清成因（锁存量） / Clear latched cause
END_IF

(* —— 段 5A：故障锁存相位迁移闸 —— *)
IF _bFault AND (_eState <> E_DL_LpiState.eFault) THEN
    _eState := E_DL_LpiState.eFault;                                     // 锁存即入故障相 / Latch enters fault phase
END_IF

(* —— 段 6：相位机（ENUM 全成员显式标签 + ELSE 兜底，R128） —— *)
CASE _eState OF

E_DL_LpiState.eIdle:
    IF _bFault THEN                                                      // 出口 1：故障锁存 / Fault latched
        _eState := E_DL_LpiState.eFault;
    ELSIF (NOT bInAuto) OR (NOT bEnable) THEN                            // 出口 2：前置不满足，明确驻留（不落 ELSE 兜底） / Precondition unmet, stay idle explicitly
        _eState := E_DL_LpiState.eIdle;
    END_IF
    (* 进相路径：段 4 阶跃检测命中时置 eCollect（进相前置与采集量重置同处一段） / Phase entry handled in segment 4 *)

E_DL_LpiState.eCollect:
    IF tonWindow.Q THEN                                                  // 出口 1：窗口到点（TON 单拍事件） / Window elapsed
        _eState := E_DL_LpiState.eEval;
    ELSIF (NOT bInAuto) OR (NOT bEnable) THEN                            // 出口 2：前置条件消失（R98 双出口） / Precondition gone
        _eState := E_DL_LpiState.eIdle;
    END_IF

E_DL_LpiState.eEval:
    fIae := LREAL_TO_REAL(_fIaeAcc);                                     // 指标定稿：IAE / Final IAE
    fIse := LREAL_TO_REAL(_fIseAcc);                                     // 指标定稿：ISE / Final ISE
    IF ABS(_fStepAmp) > DL_FLOAT_EPS THEN                                // 除零前置判 / Divide-by-zero guard
        IF _fStepAmp > 0.0 THEN
            fOvershootPct := ((_fPvPeak - fSp) / ABS(_fStepAmp)) * 100.0;   // 上行超调百分比 / Upward overshoot percentage
        ELSE
            fOvershootPct := ((fSp - _fPvPeak) / ABS(_fStepAmp)) * 100.0;   // 下行超调百分比 / Downward overshoot percentage
        END_IF
        IF fOvershootPct < 0.0 THEN
            fOvershootPct := 0.0;                                        // 无超调不报负值 / No negative overshoot
        END_IF
    ELSE
        fOvershootPct := 0.0;                                            // 阶跃量退化，超调不可算 / Degenerate step, overshoot unavailable
    END_IF
    IF _fPeakLast > DL_FLOAT_EPS THEN                                    // 除零前置判 / Divide-by-zero guard
        _fRatios := _fPeakPrev / _fPeakLast;                             // 相邻峰比 / Adjacent peak ratio
        IF _fRatios > 1.0 THEN
            fDecayRatio := 1.0;                                          // 上侧钳位 / Upper clamp
        ELSIF _fRatios < 0.0 THEN
            fDecayRatio := 0.0;                                          // 下侧钳位 / Lower clamp
        ELSE
            fDecayRatio := _fRatios;
        END_IF
    ELSE
        fDecayRatio := 0.0;                                              // 峰值不足，比值不可算 / Not enough peaks
    END_IF
    nOscCount := _nOscAcc;                                               // 振荡计数定稿 / Final oscillation count
    IF (_nOscAcc >= 4) OR (fDecayRatio > 0.60) THEN                      // 判据 1：振荡 / Criterion 1, oscillating
        eTuneHint := E_DL_LpiHint.eOscillating;
    ELSIF fOvershootPct > 20.0 THEN                                      // 判据 2：偏快 / Criterion 2, too fast
        eTuneHint := E_DL_LpiHint.eTooFast;
    ELSIF (fOvershootPct < 5.0) AND (fIae > (ABS(_fStepAmp) * DL_FLOAT_EPS)) THEN   // 判据 3：偏慢 / Criterion 3, too slow
        eTuneHint := E_DL_LpiHint.eTooSlow;
    ELSE
        eTuneHint := E_DL_LpiHint.eSuitable;                             // 默认合适 / Default suitable
    END_IF
    _uInfo := 16#0002_04B5;                                              // 信息级：本次评价完成 / Info: evaluation completed
    _eState := E_DL_LpiState.eDone;                                      // 进完成相 / Enter done phase

E_DL_LpiState.eDone:
    bEvalDone := TRUE;                                                   // 完成相保持完成位（映射到出口） / Done flag held in done phase
    IF (NOT bInAuto) OR (NOT bEnable) THEN                               // 出口 1：前置消失回空闲 / Precondition gone
        _eState := E_DL_LpiState.eIdle;
    ELSIF _bFault THEN                                                   // 出口 2：故障锁存 / Fault latched
        _eState := E_DL_LpiState.eFault;
    END_IF

E_DL_LpiState.eFault:
    ;                                                                     // 故障相：仅段 5 复位沿可迁出 / Only the reset edge leaves this phase

ELSE
    _uFault := 16#0002_03B2;                                             // 故障级：非法相位兜底（归并总码） / Illegal-phase fallback
    _bFault := TRUE;
    bError  := TRUE;
    _eCause := E_DL_LpiCause.ePhaseBad;                                  // 归因：非法相位 / Cause: illegal phase
    _eState := E_DL_LpiState.eFault;

END_CASE

(* —— 段 7：出口单点映射（名实同源；锁存码回放；故障相安全侧） —— *)
IF _bFault THEN
    bEvalDone := FALSE;                                                  // 故障相不宣称完成 / No completion claim in fault
    eTuneHint := E_DL_LpiHint.eSuitable;                                 // 故障相建议档归中性档（不外推整定建议） / Neutral hint in fault
END_IF
IF _bFault THEN
    nErrId := _uFault;                                                   // 故障锁存码回放 / Replay latched fault code
ELSE
    nErrId := _uInfo;                                                    // 信息码 / Info code
END_IF
bError := _bFault;                                                       // 故障标志与锁存同源（名实双出口，R191） / Flag from latch
eState := _eState;                                                       // 状态出口 / State outlet
eCause := _eCause;                                                       // 成因出口 / Cause outlet

END_FUNCTION_BLOCK
